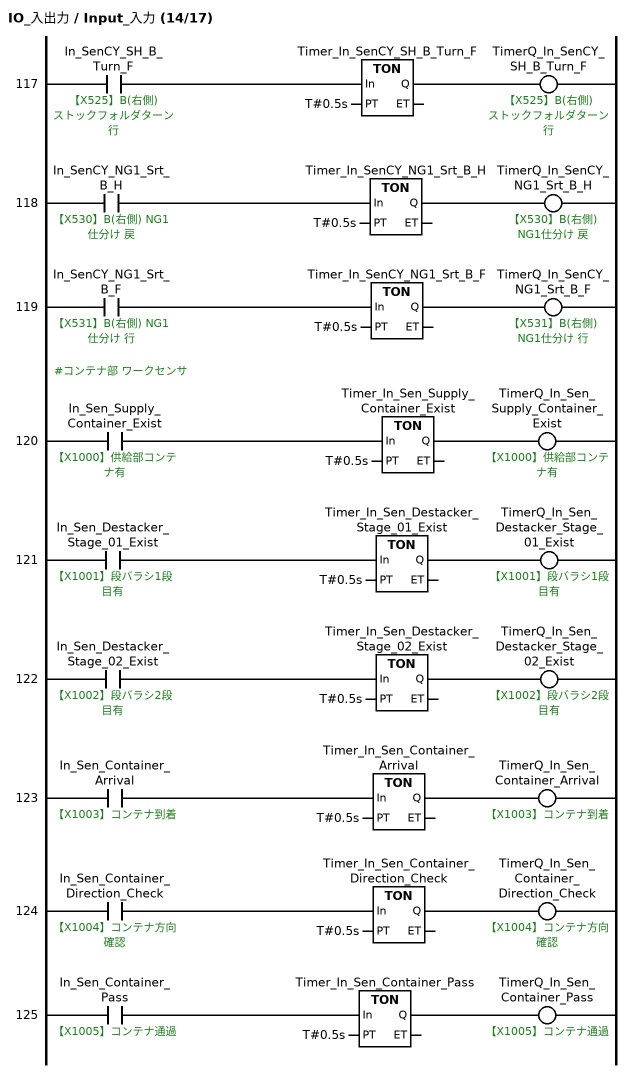
(* [picture p188: IO_入出力 / Input_入力, rungs 117-125] *)
(* Rung 117 *)
Timer_In_SenCY_SH_B_Turn_F(In := In_SenCY_SH_B_Turn_F, PT := T#0.5s);
TimerQ_In_SenCY_SH_B_Turn_F := Timer_In_SenCY_SH_B_Turn_F.Q;
(* Rung 118 *)
Timer_In_SenCY_NG1_Srt_B_H(In := In_SenCY_NG1_Srt_B_H, PT := T#0.5s);
TimerQ_In_SenCY_NG1_Srt_B_H := Timer_In_SenCY_NG1_Srt_B_H.Q;
(* Rung 119 *)
Timer_In_SenCY_NG1_Srt_B_F(In := In_SenCY_NG1_Srt_B_F, PT := T#0.5s);
TimerQ_In_SenCY_NG1_Srt_B_F := Timer_In_SenCY_NG1_Srt_B_F.Q;
(* Rung 120: #コンテナ部 ワークセンサ *)
Timer_In_Sen_Supply_Container_Exist(In := In_Sen_Supply_Container_Exist, PT := T#0.5s);
TimerQ_In_Sen_Supply_Container_Exist := Timer_In_Sen_Supply_Container_Exist.Q;
(* Rung 121 *)
Timer_In_Sen_Destacker_Stage_01_Exist(In := In_Sen_Destacker_Stage_01_Exist, PT := T#0.5s);
TimerQ_In_Sen_Destacker_Stage_01_Exist := Timer_In_Sen_Destacker_Stage_01_Exist.Q;
(* Rung 122 *)
Timer_In_Sen_Destacker_Stage_02_Exist(In := In_Sen_Destacker_Stage_02_Exist, PT := T#0.5s);
TimerQ_In_Sen_Destacker_Stage_02_Exist := Timer_In_Sen_Destacker_Stage_02_Exist.Q;
(* Rung 123 *)
Timer_In_Sen_Container_Arrival(In := In_Sen_Container_Arrival, PT := T#0.5s);
TimerQ_In_Sen_Container_Arrival := Timer_In_Sen_Container_Arrival.Q;
(* Rung 124 *)
Timer_In_Sen_Container_Direction_Check(In := In_Sen_Container_Direction_Check, PT := T#0.5s);
TimerQ_In_Sen_Container_Direction_Check := Timer_In_Sen_Container_Direction_Check.Q;
(* Rung 125 *)
Timer_In_Sen_Container_Pass(In := In_Sen_Container_Pass, PT := T#0.5s);
TimerQ_In_Sen_Container_Pass := Timer_In_Sen_Container_Pass.Q;

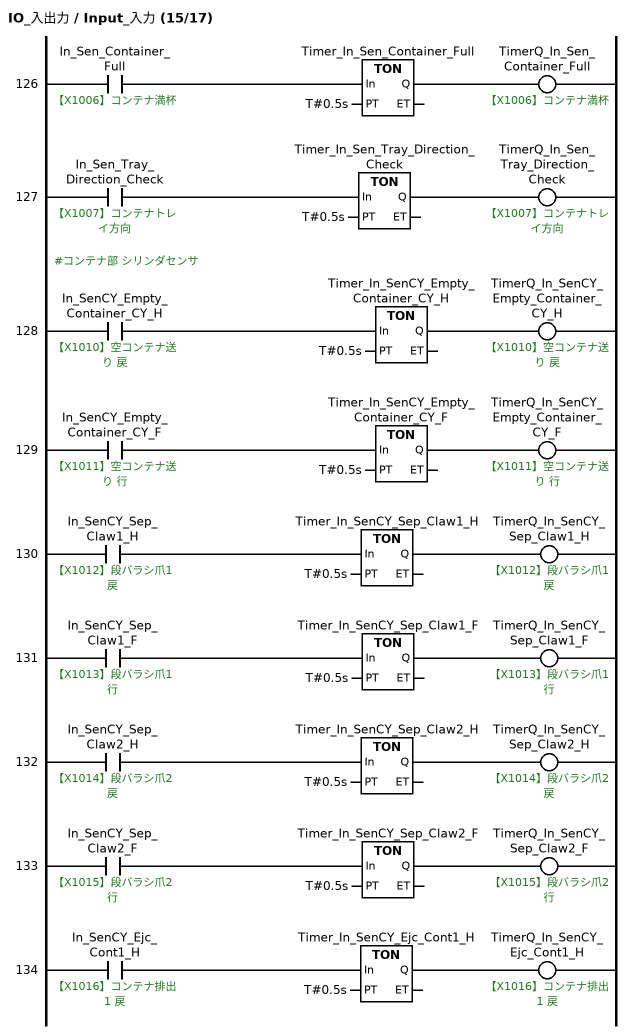
(* Rung 126 *)
Timer_In_Sen_Container_Full(In := In_Sen_Container_Full, PT := T#0.5s);
TimerQ_In_Sen_Container_Full := Timer_In_Sen_Container_Full.Q;
(* Rung 127 *)
Timer_In_Sen_Tray_Direction_Check(In := In_Sen_Tray_Direction_Check, PT := T#0.5s);
TimerQ_In_Sen_Tray_Direction_Check := Timer_In_Sen_Tray_Direction_Check.Q;
(* Rung 128: #コンテナ部 シリンダセンサ *)
Timer_In_SenCY_Empty_Container_CY_H(In := In_SenCY_Empty_Container_CY_H, PT := T#0.5s);
TimerQ_In_SenCY_Empty_Container_CY_H := Timer_In_SenCY_Empty_Container_CY_H.Q;
(* Rung 129 *)
Timer_In_SenCY_Empty_Container_CY_F(In := In_SenCY_Empty_Container_CY_F, PT := T#0.5s);
TimerQ_In_SenCY_Empty_Container_CY_F := Timer_In_SenCY_Empty_Container_CY_F.Q;
(* Rung 130 *)
Timer_In_SenCY_Sep_Claw1_H(In := In_SenCY_Sep_Claw1_H, PT := T#0.5s);
TimerQ_In_SenCY_Sep_Claw1_H := Timer_In_SenCY_Sep_Claw1_H.Q;
(* Rung 131 *)
Timer_In_SenCY_Sep_Claw1_F(In := In_SenCY_Sep_Claw1_F, PT := T#0.5s);
TimerQ_In_SenCY_Sep_Claw1_F := Timer_In_SenCY_Sep_Claw1_F.Q;
(* Rung 132 *)
Timer_In_SenCY_Sep_Claw2_H(In := In_SenCY_Sep_Claw2_H, PT := T#0.5s);
TimerQ_In_SenCY_Sep_Claw2_H := Timer_In_SenCY_Sep_Claw2_H.Q;
(* Rung 133 *)
Timer_In_SenCY_Sep_Claw2_F(In := In_SenCY_Sep_Claw2_F, PT := T#0.5s);
TimerQ_In_SenCY_Sep_Claw2_F := Timer_In_SenCY_Sep_Claw2_F.Q;
(* Rung 134 *)
Timer_In_SenCY_Ejc_Cont1_H(In := In_SenCY_Ejc_Cont1_H, PT := T#0.5s);
TimerQ_In_SenCY_Ejc_Cont1_H := Timer_In_SenCY_Ejc_Cont1_H.Q;

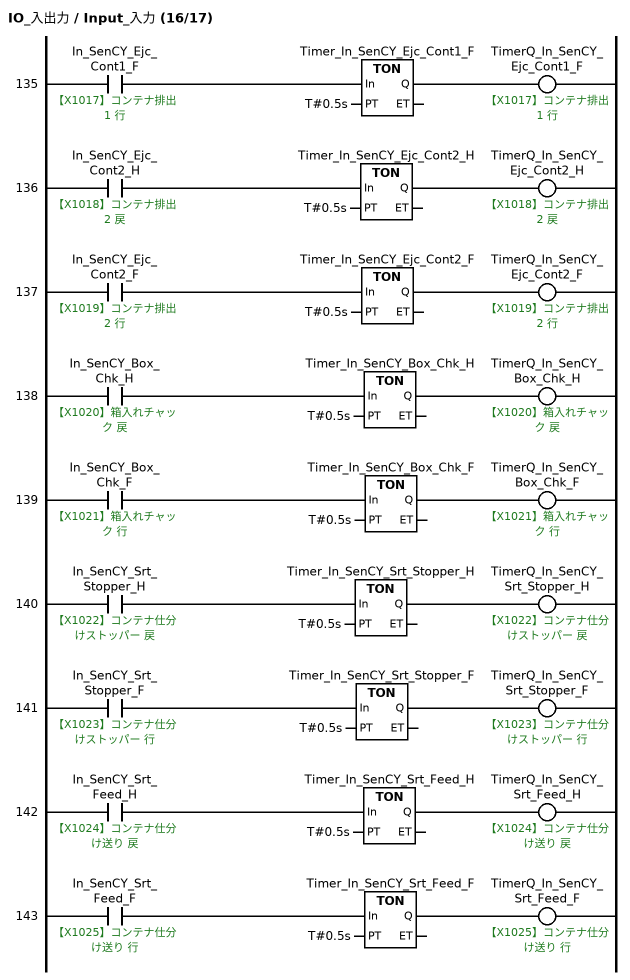
(* Rung 135 *)
Timer_In_SenCY_Ejc_Cont1_F(In := In_SenCY_Ejc_Cont1_F, PT := T#0.5s);
TimerQ_In_SenCY_Ejc_Cont1_F := Timer_In_SenCY_Ejc_Cont1_F.Q;
(* Rung 136 *)
Timer_In_SenCY_Ejc_Cont2_H(In := In_SenCY_Ejc_Cont2_H, PT := T#0.5s);
TimerQ_In_SenCY_Ejc_Cont2_H := Timer_In_SenCY_Ejc_Cont2_H.Q;
(* Rung 137 *)
Timer_In_SenCY_Ejc_Cont2_F(In := In_SenCY_Ejc_Cont2_F, PT := T#0.5s);
TimerQ_In_SenCY_Ejc_Cont2_F := Timer_In_SenCY_Ejc_Cont2_F.Q;
(* Rung 138 *)
Timer_In_SenCY_Box_Chk_H(In := In_SenCY_Box_Chk_H, PT := T#0.5s);
TimerQ_In_SenCY_Box_Chk_H := Timer_In_SenCY_Box_Chk_H.Q;
(* Rung 139 *)
Timer_In_SenCY_Box_Chk_F(In := In_SenCY_Box_Chk_F, PT := T#0.5s);
TimerQ_In_SenCY_Box_Chk_F := Timer_In_SenCY_Box_Chk_F.Q;
(* Rung 140 *)
Timer_In_SenCY_Srt_Stopper_H(In := In_SenCY_Srt_Stopper_H, PT := T#0.5s);
TimerQ_In_SenCY_Srt_Stopper_H := Timer_In_SenCY_Srt_Stopper_H.Q;
(* Rung 141 *)
Timer_In_SenCY_Srt_Stopper_F(In := In_SenCY_Srt_Stopper_F, PT := T#0.5s);
TimerQ_In_SenCY_Srt_Stopper_F := Timer_In_SenCY_Srt_Stopper_F.Q;
(* Rung 142 *)
Timer_In_SenCY_Srt_Feed_H(In := In_SenCY_Srt_Feed_H, PT := T#0.5s);
TimerQ_In_SenCY_Srt_Feed_H := Timer_In_SenCY_Srt_Feed_H.Q;
(* Rung 143 *)
Timer_In_SenCY_Srt_Feed_F(In := In_SenCY_Srt_Feed_F, PT := T#0.5s);
TimerQ_In_SenCY_Srt_Feed_F := Timer_In_SenCY_Srt_Feed_F.Q;

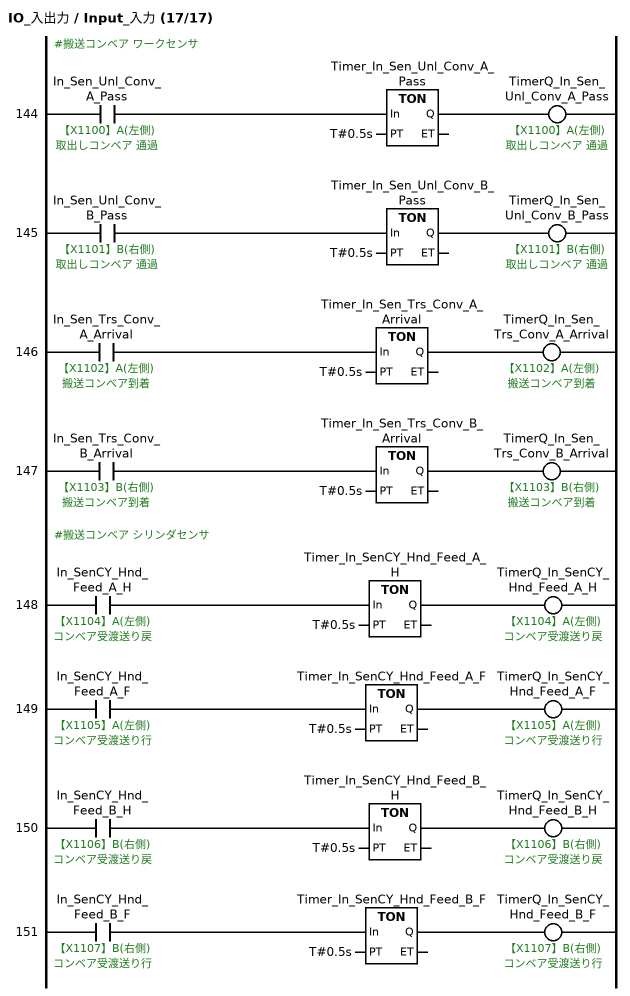
(* Rung 144: #搬送コンベア ワークセンサ *)
Timer_In_Sen_Unl_Conv_A_Pass(In := In_Sen_Unl_Conv_A_Pass, PT := T#0.5s);
TimerQ_In_Sen_Unl_Conv_A_Pass := Timer_In_Sen_Unl_Conv_A_Pass.Q;
(* Rung 145 *)
Timer_In_Sen_Unl_Conv_B_Pass(In := In_Sen_Unl_Conv_B_Pass, PT := T#0.5s);
TimerQ_In_Sen_Unl_Conv_B_Pass := Timer_In_Sen_Unl_Conv_B_Pass.Q;
(* Rung 146 *)
Timer_In_Sen_Trs_Conv_A_Arrival(In := In_Sen_Trs_Conv_A_Arrival, PT := T#0.5s);
TimerQ_In_Sen_Trs_Conv_A_Arrival := Timer_In_Sen_Trs_Conv_A_Arrival.Q;
(* Rung 147 *)
Timer_In_Sen_Trs_Conv_B_Arrival(In := In_Sen_Trs_Conv_B_Arrival, PT := T#0.5s);
TimerQ_In_Sen_Trs_Conv_B_Arrival := Timer_In_Sen_Trs_Conv_B_Arrival.Q;
(* Rung 148: #搬送コンベア シリンダセンサ *)
Timer_In_SenCY_Hnd_Feed_A_H(In := In_SenCY_Hnd_Feed_A_H, PT := T#0.5s);
TimerQ_In_SenCY_Hnd_Feed_A_H := Timer_In_SenCY_Hnd_Feed_A_H.Q;
(* Rung 149 *)
Timer_In_SenCY_Hnd_Feed_A_F(In := In_SenCY_Hnd_Feed_A_F, PT := T#0.5s);
TimerQ_In_SenCY_Hnd_Feed_A_F := Timer_In_SenCY_Hnd_Feed_A_F.Q;
(* Rung 150 *)
Timer_In_SenCY_Hnd_Feed_B_H(In := In_SenCY_Hnd_Feed_B_H, PT := T#0.5s);
TimerQ_In_SenCY_Hnd_Feed_B_H := Timer_In_SenCY_Hnd_Feed_B_H.Q;
(* Rung 151 *)
Timer_In_SenCY_Hnd_Feed_B_F(In := In_SenCY_Hnd_Feed_B_F, PT := T#0.5s);
TimerQ_In_SenCY_Hnd_Feed_B_F := Timer_In_SenCY_Hnd_Feed_B_F.Q;

(* Section Output_出力: ladder, written here as Structured Text *)

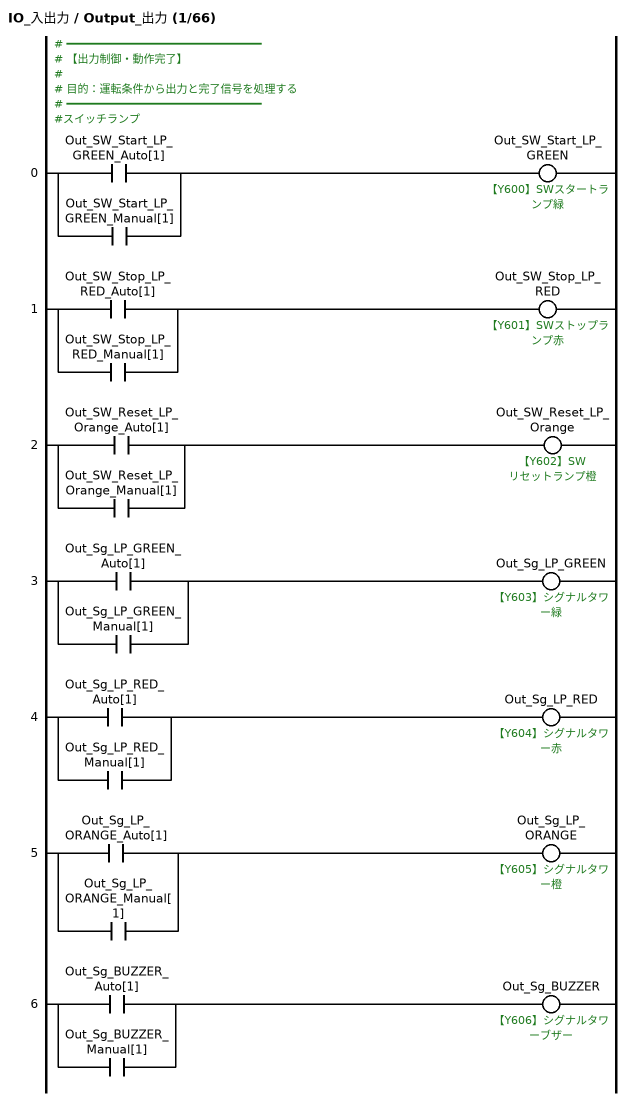
(* Rung 0: # ━━━━━━━━━━━━━━━━━━━━━━━━━━━━━━ / # 【出力制御・動作完了】 / # / # 目的：運転条件から出力と完了信号を処理する / # ━━━━━━━━━━━━━━━━━━━━━━━━━━━━━━ / #スイッチランプ *)
Out_SW_Start_LP_GREEN := Out_SW_Start_LP_GREEN_Auto[1] OR Out_SW_Start_LP_GREEN_Manual[1];
(* Rung 1 *)
Out_SW_Stop_LP_RED := Out_SW_Stop_LP_RED_Auto[1] OR Out_SW_Stop_LP_RED_Manual[1];
(* Rung 2 *)
Out_SW_Reset_LP_Orange := Out_SW_Reset_LP_Orange_Auto[1] OR Out_SW_Reset_LP_Orange_Manual[1];
(* Rung 3 *)
Out_Sg_LP_GREEN := Out_Sg_LP_GREEN_Auto[1] OR Out_Sg_LP_GREEN_Manual[1];
(* Rung 4 *)
Out_Sg_LP_RED := Out_Sg_LP_RED_Auto[1] OR Out_Sg_LP_RED_Manual[1];
(* Rung 5 *)
Out_Sg_LP_ORANGE := Out_Sg_LP_ORANGE_Auto[1] OR Out_Sg_LP_ORANGE_Manual[1];
(* Rung 6 *)
Out_Sg_BUZZER := Out_Sg_BUZZER_Auto[1] OR Out_Sg_BUZZER_Manual[1];

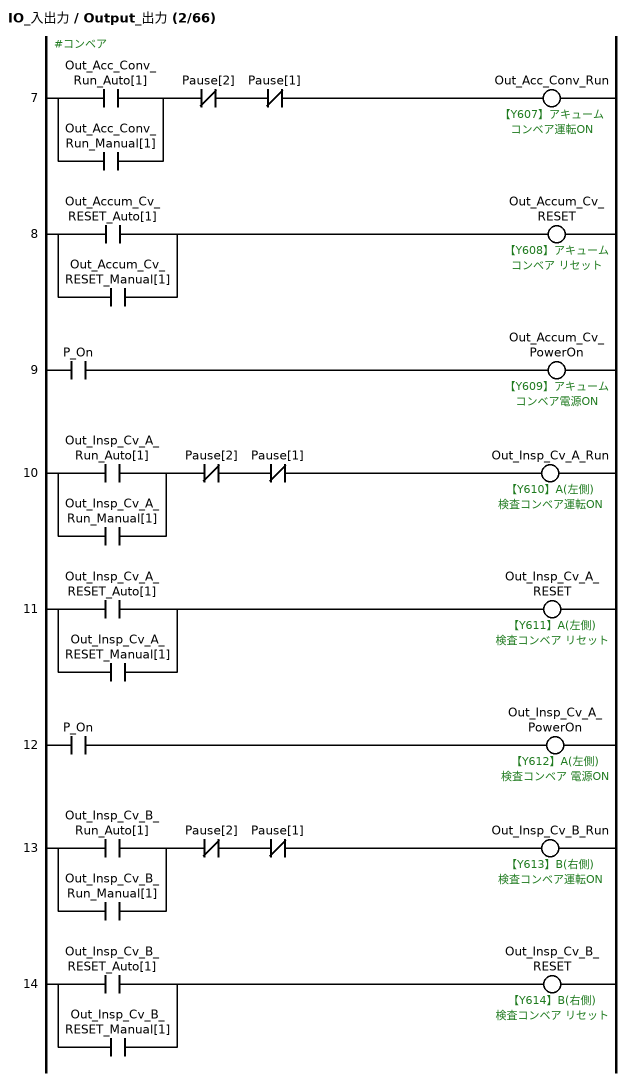
(* Rung 7: #コンベア *)
Out_Acc_Conv_Run := (Out_Acc_Conv_Run_Auto[1] OR Out_Acc_Conv_Run_Manual[1]) AND NOT Pause[2] AND NOT Pause[1];
(* Rung 8 *)
Out_Accum_Cv_RESET := Out_Accum_Cv_RESET_Auto[1] OR Out_Accum_Cv_RESET_Manual[1];
(* Rung 9 *)
Out_Accum_Cv_PowerOn := P_On;
(* Rung 10 *)
Out_Insp_Cv_A_Run := (Out_Insp_Cv_A_Run_Auto[1] OR Out_Insp_Cv_A_Run_Manual[1]) AND NOT Pause[2] AND NOT Pause[1];
(* Rung 11 *)
Out_Insp_Cv_A_RESET := Out_Insp_Cv_A_RESET_Auto[1] OR Out_Insp_Cv_A_RESET_Manual[1];
(* Rung 12 *)
Out_Insp_Cv_A_PowerOn := P_On;
(* Rung 13 *)
Out_Insp_Cv_B_Run := (Out_Insp_Cv_B_Run_Auto[1] OR Out_Insp_Cv_B_Run_Manual[1]) AND NOT Pause[2] AND NOT Pause[1];
(* Rung 14 *)
Out_Insp_Cv_B_RESET := Out_Insp_Cv_B_RESET_Auto[1] OR Out_Insp_Cv_B_RESET_Manual[1];

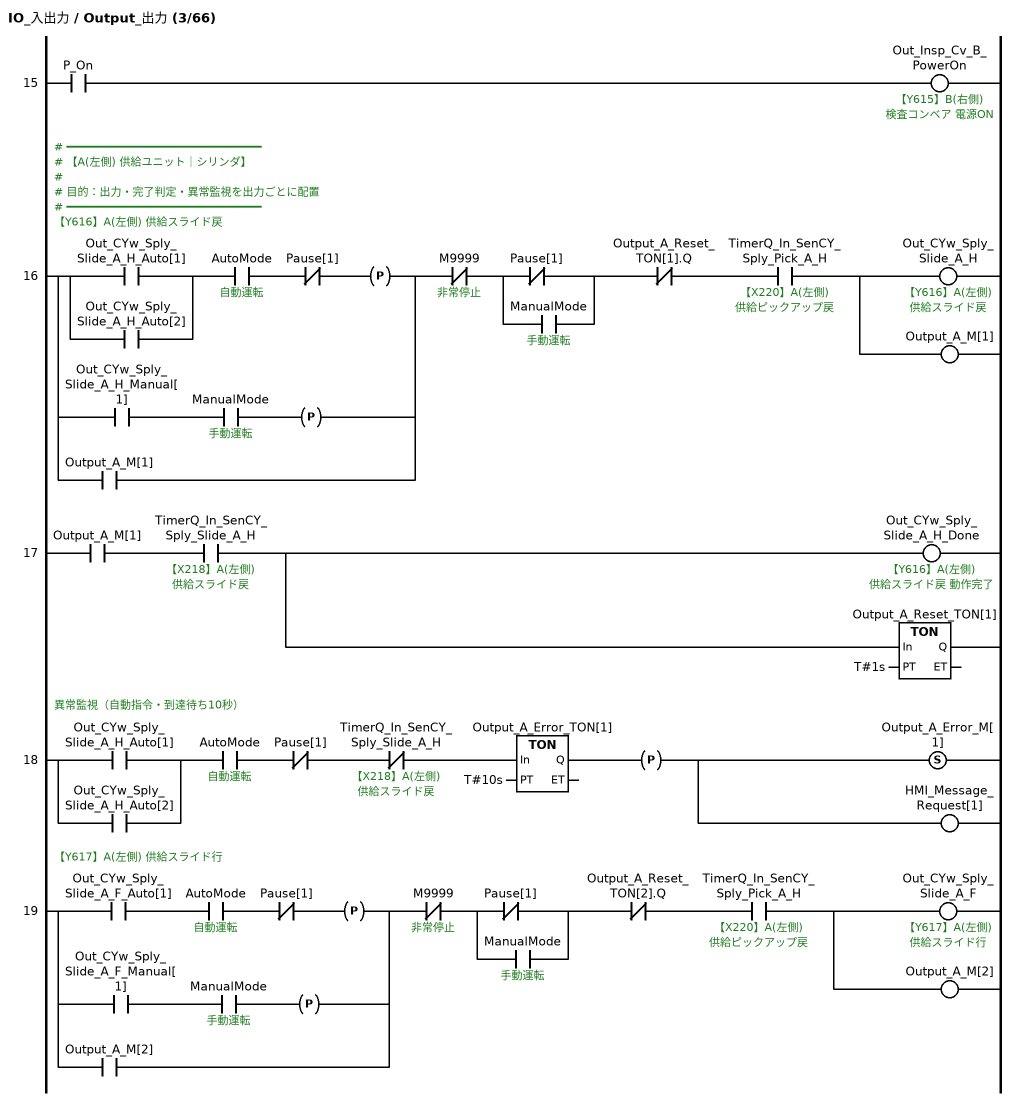
(* Rung 15 *)
Out_Insp_Cv_B_PowerOn := P_On;
(* Rung 16: # ━━━━━━━━━━━━━━━━━━━━━━━━━━━━━━ / # 【A(左側) 供給ユニット｜シリンダ】 / # / # 目的：出力・完了判定・異常監視を出力ごとに配置 / # ━━━━━━━━━━━━━━━━━━━━━━━━━━━━━━ / 【Y616】A(左側) 供給スライド戻 *)
_e1(CLK := (Out_CYw_Sply_Slide_A_H_Auto[1] OR Out_CYw_Sply_Slide_A_H_Auto[2]) AND AutoMode AND NOT Pause[1]);
_e2(CLK := Out_CYw_Sply_Slide_A_H_Manual[1] AND ManualMode);
_p3 := (_e1.Q OR _e2.Q OR Output_A_M[1]) AND NOT M9999 AND (NOT Pause[1] OR ManualMode) AND NOT Output_A_Reset_TON[1].Q AND TimerQ_In_SenCY_Sply_Pick_A_H;
Out_CYw_Sply_Slide_A_H := _p3;
Output_A_M[1] := _p3;
(* Rung 17 *)
Out_CYw_Sply_Slide_A_H_Done := Output_A_M[1] AND TimerQ_In_SenCY_Sply_Slide_A_H;
Output_A_Reset_TON[1](In := Output_A_M[1] AND TimerQ_In_SenCY_Sply_Slide_A_H, PT := T#1s);
(* Rung 18: 異常監視（自動指令・到達待ち10秒） *)
Output_A_Error_TON[1](In := (Out_CYw_Sply_Slide_A_H_Auto[1] OR Out_CYw_Sply_Slide_A_H_Auto[2]) AND AutoMode AND NOT Pause[1] AND NOT TimerQ_In_SenCY_Sply_Slide_A_H, PT := T#10s);
_e4(CLK := Output_A_Error_TON[1].Q);
IF _e4.Q THEN Output_A_Error_M[1] := TRUE; END_IF;
HMI_Message_Request[1] := _e4.Q;
(* Rung 19: 【Y617】A(左側) 供給スライド行 *)
_e5(CLK := Out_CYw_Sply_Slide_A_F_Auto[1] AND AutoMode AND NOT Pause[1]);
_e6(CLK := Out_CYw_Sply_Slide_A_F_Manual[1] AND ManualMode);
_p7 := (_e5.Q OR _e6.Q OR Output_A_M[2]) AND NOT M9999 AND (NOT Pause[1] OR ManualMode) AND NOT Output_A_Reset_TON[2].Q AND TimerQ_In_SenCY_Sply_Pick_A_H;
Out_CYw_Sply_Slide_A_F := _p7;
Output_A_M[2] := _p7;

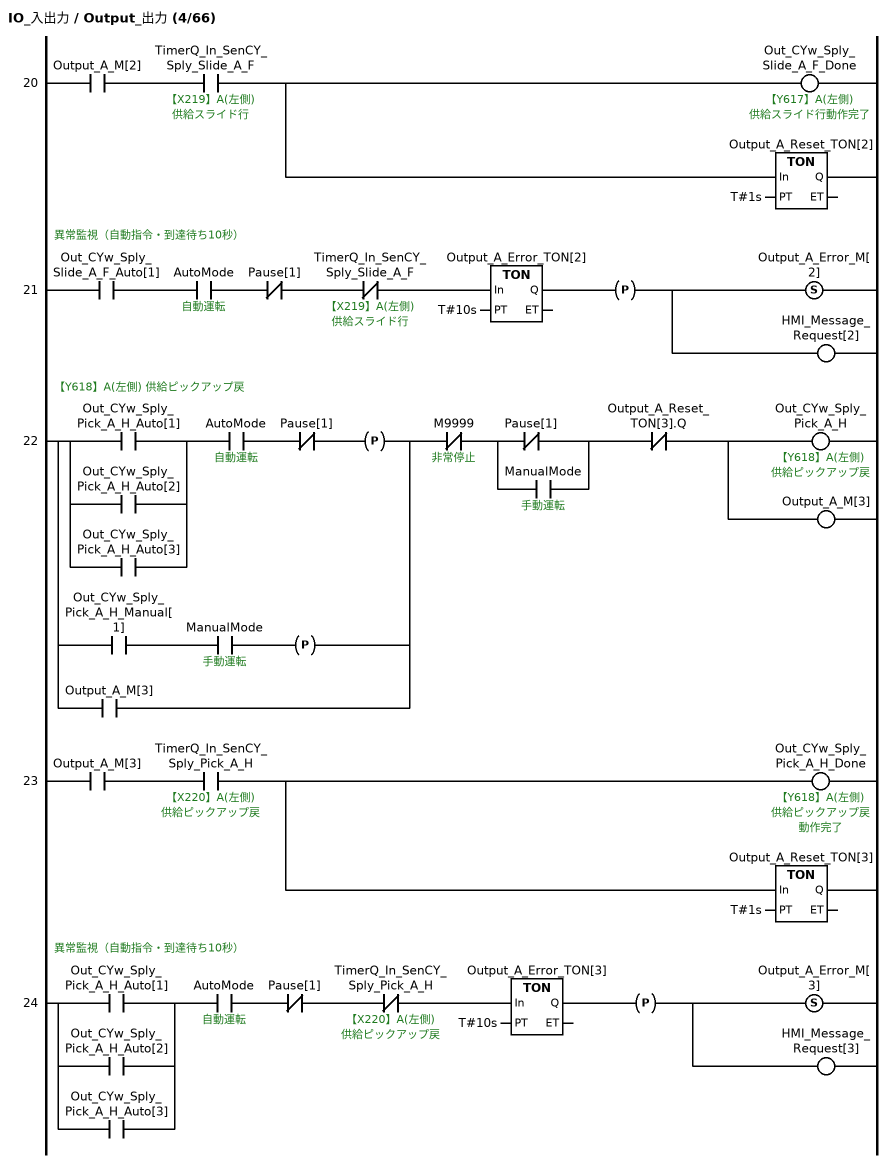
(* Rung 20 *)
Out_CYw_Sply_Slide_A_F_Done := Output_A_M[2] AND TimerQ_In_SenCY_Sply_Slide_A_F;
Output_A_Reset_TON[2](In := Output_A_M[2] AND TimerQ_In_SenCY_Sply_Slide_A_F, PT := T#1s);
(* Rung 21: 異常監視（自動指令・到達待ち10秒） *)
Output_A_Error_TON[2](In := Out_CYw_Sply_Slide_A_F_Auto[1] AND AutoMode AND NOT Pause[1] AND NOT TimerQ_In_SenCY_Sply_Slide_A_F, PT := T#10s);
_e8(CLK := Output_A_Error_TON[2].Q);
IF _e8.Q THEN Output_A_Error_M[2] := TRUE; END_IF;
HMI_Message_Request[2] := _e8.Q;
(* Rung 22: 【Y618】A(左側) 供給ピックアップ戻 *)
_e9(CLK := (Out_CYw_Sply_Pick_A_H_Auto[1] OR Out_CYw_Sply_Pick_A_H_Auto[2] OR Out_CYw_Sply_Pick_A_H_Auto[3]) AND AutoMode AND NOT Pause[1]);
_e10(CLK := Out_CYw_Sply_Pick_A_H_Manual[1] AND ManualMode);
_p11 := (_e9.Q OR _e10.Q OR Output_A_M[3]) AND NOT M9999 AND (NOT Pause[1] OR ManualMode) AND NOT Output_A_Reset_TON[3].Q;
Out_CYw_Sply_Pick_A_H := _p11;
Output_A_M[3] := _p11;
(* Rung 23 *)
Out_CYw_Sply_Pick_A_H_Done := Output_A_M[3] AND TimerQ_In_SenCY_Sply_Pick_A_H;
Output_A_Reset_TON[3](In := Output_A_M[3] AND TimerQ_In_SenCY_Sply_Pick_A_H, PT := T#1s);
(* Rung 24: 異常監視（自動指令・到達待ち10秒） *)
Output_A_Error_TON[3](In := (Out_CYw_Sply_Pick_A_H_Auto[1] OR Out_CYw_Sply_Pick_A_H_Auto[2] OR Out_CYw_Sply_Pick_A_H_Auto[3]) AND AutoMode AND NOT Pause[1] AND NOT TimerQ_In_SenCY_Sply_Pick_A_H, PT := T#10s);
_e12(CLK := Output_A_Error_TON[3].Q);
IF _e12.Q THEN Output_A_Error_M[3] := TRUE; END_IF;
HMI_Message_Request[3] := _e12.Q;

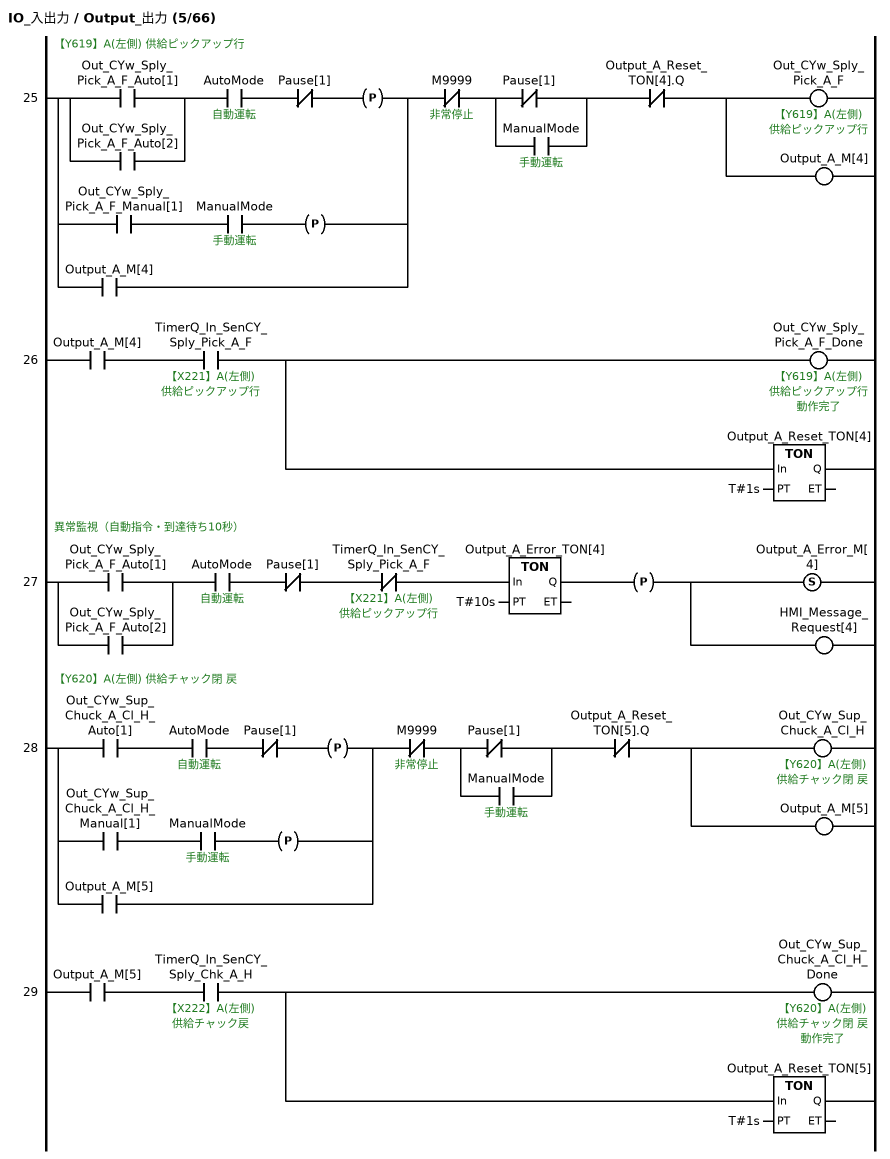
(* Rung 25: 【Y619】A(左側) 供給ピックアップ行 *)
_e13(CLK := (Out_CYw_Sply_Pick_A_F_Auto[1] OR Out_CYw_Sply_Pick_A_F_Auto[2]) AND AutoMode AND NOT Pause[1]);
_e14(CLK := Out_CYw_Sply_Pick_A_F_Manual[1] AND ManualMode);
_p15 := (_e13.Q OR _e14.Q OR Output_A_M[4]) AND NOT M9999 AND (NOT Pause[1] OR ManualMode) AND NOT Output_A_Reset_TON[4].Q;
Out_CYw_Sply_Pick_A_F := _p15;
Output_A_M[4] := _p15;
(* Rung 26 *)
Out_CYw_Sply_Pick_A_F_Done := Output_A_M[4] AND TimerQ_In_SenCY_Sply_Pick_A_F;
Output_A_Reset_TON[4](In := Output_A_M[4] AND TimerQ_In_SenCY_Sply_Pick_A_F, PT := T#1s);
(* Rung 27: 異常監視（自動指令・到達待ち10秒） *)
Output_A_Error_TON[4](In := (Out_CYw_Sply_Pick_A_F_Auto[1] OR Out_CYw_Sply_Pick_A_F_Auto[2]) AND AutoMode AND NOT Pause[1] AND NOT TimerQ_In_SenCY_Sply_Pick_A_F, PT := T#10s);
_e16(CLK := Output_A_Error_TON[4].Q);
IF _e16.Q THEN Output_A_Error_M[4] := TRUE; END_IF;
HMI_Message_Request[4] := _e16.Q;
(* Rung 28: 【Y620】A(左側) 供給チャック閉 戻 *)
_e17(CLK := Out_CYw_Sup_Chuck_A_Cl_H_Auto[1] AND AutoMode AND NOT Pause[1]);
_e18(CLK := Out_CYw_Sup_Chuck_A_Cl_H_Manual[1] AND ManualMode);
_p19 := (_e17.Q OR _e18.Q OR Output_A_M[5]) AND NOT M9999 AND (NOT Pause[1] OR ManualMode) AND NOT Output_A_Reset_TON[5].Q;
Out_CYw_Sup_Chuck_A_Cl_H := _p19;
Output_A_M[5] := _p19;
(* Rung 29 *)
Out_CYw_Sup_Chuck_A_Cl_H_Done := Output_A_M[5] AND TimerQ_In_SenCY_Sply_Chk_A_H;
Output_A_Reset_TON[5](In := Output_A_M[5] AND TimerQ_In_SenCY_Sply_Chk_A_H, PT := T#1s);

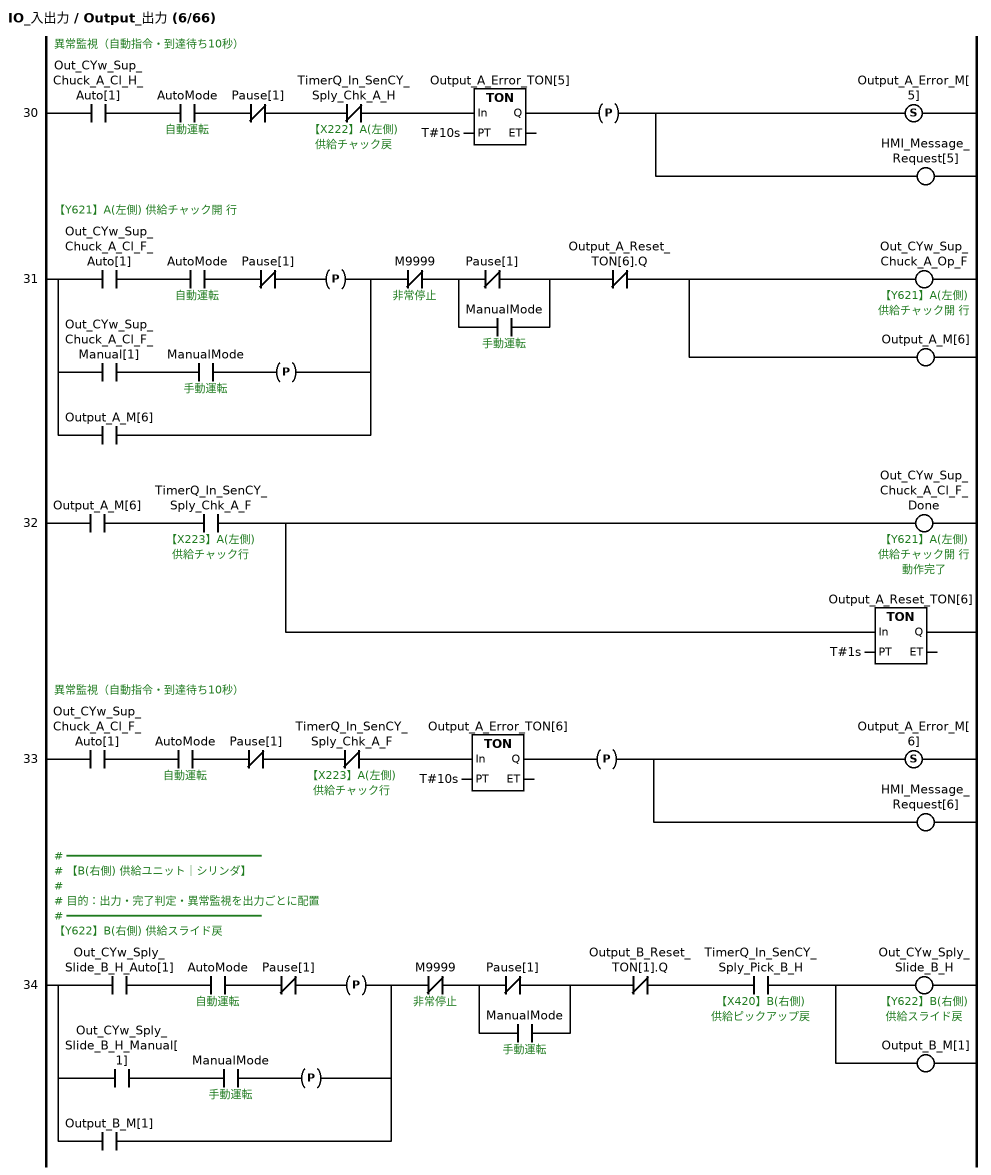
(* Rung 30: 異常監視（自動指令・到達待ち10秒） *)
Output_A_Error_TON[5](In := Out_CYw_Sup_Chuck_A_Cl_H_Auto[1] AND AutoMode AND NOT Pause[1] AND NOT TimerQ_In_SenCY_Sply_Chk_A_H, PT := T#10s);
_e20(CLK := Output_A_Error_TON[5].Q);
IF _e20.Q THEN Output_A_Error_M[5] := TRUE; END_IF;
HMI_Message_Request[5] := _e20.Q;
(* Rung 31: 【Y621】A(左側) 供給チャック開 行 *)
_e21(CLK := Out_CYw_Sup_Chuck_A_Cl_F_Auto[1] AND AutoMode AND NOT Pause[1]);
_e22(CLK := Out_CYw_Sup_Chuck_A_Cl_F_Manual[1] AND ManualMode);
_p23 := (_e21.Q OR _e22.Q OR Output_A_M[6]) AND NOT M9999 AND (NOT Pause[1] OR ManualMode) AND NOT Output_A_Reset_TON[6].Q;
Out_CYw_Sup_Chuck_A_Op_F := _p23;
Output_A_M[6] := _p23;
(* Rung 32 *)
Out_CYw_Sup_Chuck_A_Cl_F_Done := Output_A_M[6] AND TimerQ_In_SenCY_Sply_Chk_A_F;
Output_A_Reset_TON[6](In := Output_A_M[6] AND TimerQ_In_SenCY_Sply_Chk_A_F, PT := T#1s);
(* Rung 33: 異常監視（自動指令・到達待ち10秒） *)
Output_A_Error_TON[6](In := Out_CYw_Sup_Chuck_A_Cl_F_Auto[1] AND AutoMode AND NOT Pause[1] AND NOT TimerQ_In_SenCY_Sply_Chk_A_F, PT := T#10s);
_e24(CLK := Output_A_Error_TON[6].Q);
IF _e24.Q THEN Output_A_Error_M[6] := TRUE; END_IF;
HMI_Message_Request[6] := _e24.Q;
(* Rung 34: # ━━━━━━━━━━━━━━━━━━━━━━━━━━━━━━ / # 【B(右側) 供給ユニット｜シリンダ】 / # / # 目的：出力・完了判定・異常監視を出力ごとに配置 / # ━━━━━━━━━━━━━━━━━━━━━━━━━━━━━━ / 【Y622】B(右側) 供給スライド戻 *)
_e25(CLK := Out_CYw_Sply_Slide_B_H_Auto[1] AND AutoMode AND NOT Pause[1]);
_e26(CLK := Out_CYw_Sply_Slide_B_H_Manual[1] AND ManualMode);
_p27 := (_e25.Q OR _e26.Q OR Output_B_M[1]) AND NOT M9999 AND (NOT Pause[1] OR ManualMode) AND NOT Output_B_Reset_TON[1].Q AND TimerQ_In_SenCY_Sply_Pick_B_H;
Out_CYw_Sply_Slide_B_H := _p27;
Output_B_M[1] := _p27;

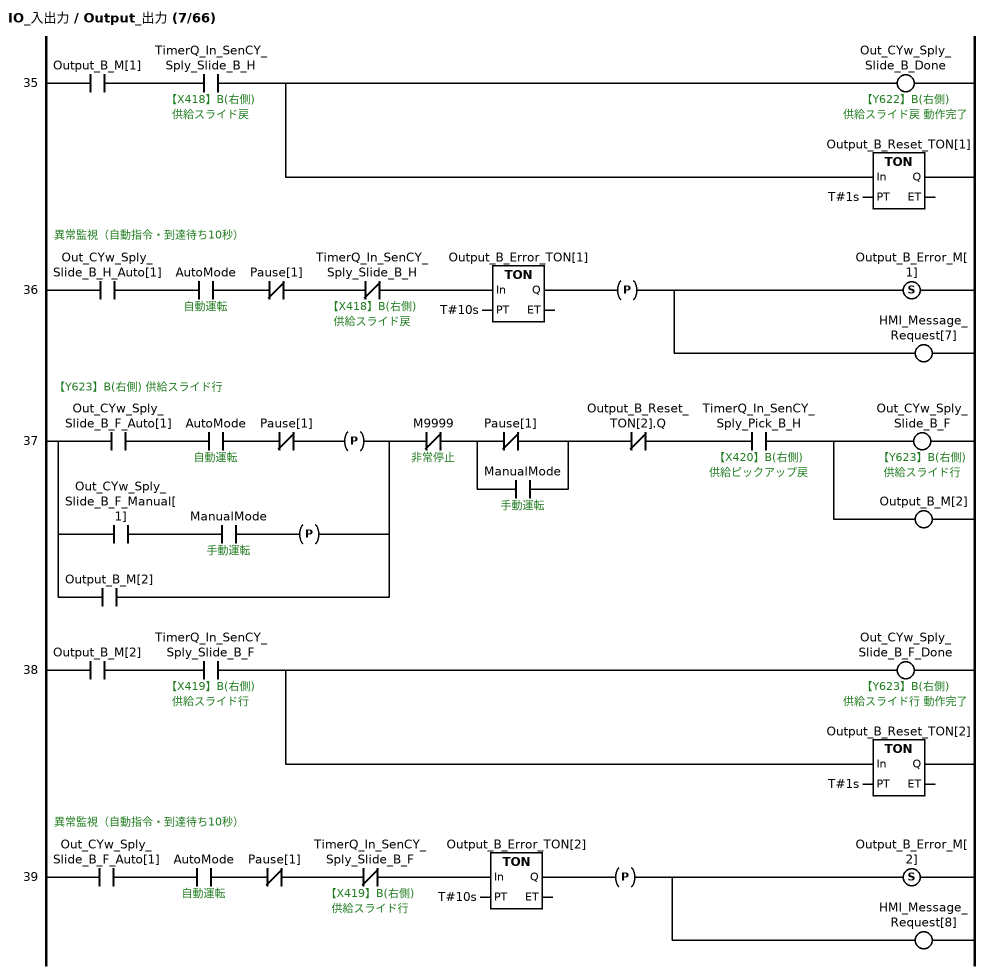
(* Rung 35 *)
Out_CYw_Sply_Slide_B_Done := Output_B_M[1] AND TimerQ_In_SenCY_Sply_Slide_B_H;
Output_B_Reset_TON[1](In := Output_B_M[1] AND TimerQ_In_SenCY_Sply_Slide_B_H, PT := T#1s);
(* Rung 36: 異常監視（自動指令・到達待ち10秒） *)
Output_B_Error_TON[1](In := Out_CYw_Sply_Slide_B_H_Auto[1] AND AutoMode AND NOT Pause[1] AND NOT TimerQ_In_SenCY_Sply_Slide_B_H, PT := T#10s);
_e28(CLK := Output_B_Error_TON[1].Q);
IF _e28.Q THEN Output_B_Error_M[1] := TRUE; END_IF;
HMI_Message_Request[7] := _e28.Q;
(* Rung 37: 【Y623】B(右側) 供給スライド行 *)
_e29(CLK := Out_CYw_Sply_Slide_B_F_Auto[1] AND AutoMode AND NOT Pause[1]);
_e30(CLK := Out_CYw_Sply_Slide_B_F_Manual[1] AND ManualMode);
_p31 := (_e29.Q OR _e30.Q OR Output_B_M[2]) AND NOT M9999 AND (NOT Pause[1] OR ManualMode) AND NOT Output_B_Reset_TON[2].Q AND TimerQ_In_SenCY_Sply_Pick_B_H;
Out_CYw_Sply_Slide_B_F := _p31;
Output_B_M[2] := _p31;
(* Rung 38 *)
Out_CYw_Sply_Slide_B_F_Done := Output_B_M[2] AND TimerQ_In_SenCY_Sply_Slide_B_F;
Output_B_Reset_TON[2](In := Output_B_M[2] AND TimerQ_In_SenCY_Sply_Slide_B_F, PT := T#1s);
(* Rung 39: 異常監視（自動指令・到達待ち10秒） *)
Output_B_Error_TON[2](In := Out_CYw_Sply_Slide_B_F_Auto[1] AND AutoMode AND NOT Pause[1] AND NOT TimerQ_In_SenCY_Sply_Slide_B_F, PT := T#10s);
_e32(CLK := Output_B_Error_TON[2].Q);
IF _e32.Q THEN Output_B_Error_M[2] := TRUE; END_IF;
HMI_Message_Request[8] := _e32.Q;

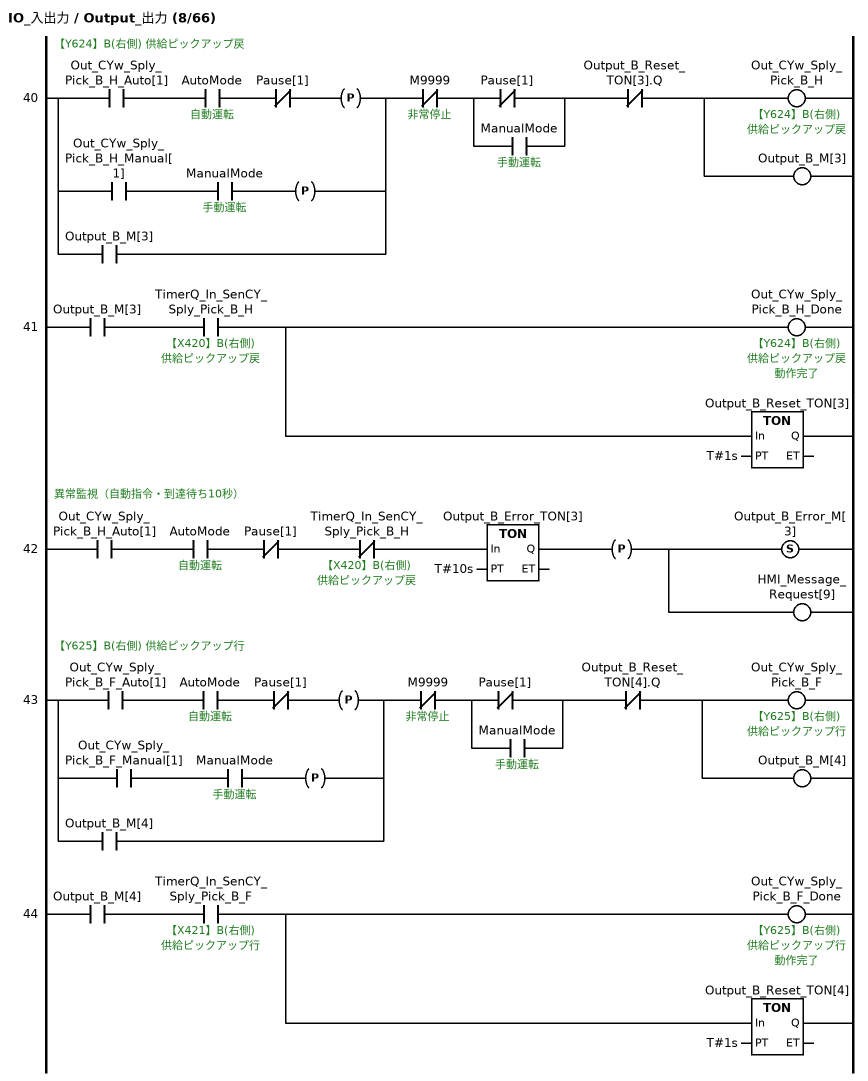
(* Rung 40: 【Y624】B(右側) 供給ピックアップ戻 *)
_e33(CLK := Out_CYw_Sply_Pick_B_H_Auto[1] AND AutoMode AND NOT Pause[1]);
_e34(CLK := Out_CYw_Sply_Pick_B_H_Manual[1] AND ManualMode);
_p35 := (_e33.Q OR _e34.Q OR Output_B_M[3]) AND NOT M9999 AND (NOT Pause[1] OR ManualMode) AND NOT Output_B_Reset_TON[3].Q;
Out_CYw_Sply_Pick_B_H := _p35;
Output_B_M[3] := _p35;
(* Rung 41 *)
Out_CYw_Sply_Pick_B_H_Done := Output_B_M[3] AND TimerQ_In_SenCY_Sply_Pick_B_H;
Output_B_Reset_TON[3](In := Output_B_M[3] AND TimerQ_In_SenCY_Sply_Pick_B_H, PT := T#1s);
(* Rung 42: 異常監視（自動指令・到達待ち10秒） *)
Output_B_Error_TON[3](In := Out_CYw_Sply_Pick_B_H_Auto[1] AND AutoMode AND NOT Pause[1] AND NOT TimerQ_In_SenCY_Sply_Pick_B_H, PT := T#10s);
_e36(CLK := Output_B_Error_TON[3].Q);
IF _e36.Q THEN Output_B_Error_M[3] := TRUE; END_IF;
HMI_Message_Request[9] := _e36.Q;
(* Rung 43: 【Y625】B(右側) 供給ピックアップ行 *)
_e37(CLK := Out_CYw_Sply_Pick_B_F_Auto[1] AND AutoMode AND NOT Pause[1]);
_e38(CLK := Out_CYw_Sply_Pick_B_F_Manual[1] AND ManualMode);
_p39 := (_e37.Q OR _e38.Q OR Output_B_M[4]) AND NOT M9999 AND (NOT Pause[1] OR ManualMode) AND NOT Output_B_Reset_TON[4].Q;
Out_CYw_Sply_Pick_B_F := _p39;
Output_B_M[4] := _p39;
(* Rung 44 *)
Out_CYw_Sply_Pick_B_F_Done := Output_B_M[4] AND TimerQ_In_SenCY_Sply_Pick_B_F;
Output_B_Reset_TON[4](In := Output_B_M[4] AND TimerQ_In_SenCY_Sply_Pick_B_F, PT := T#1s);

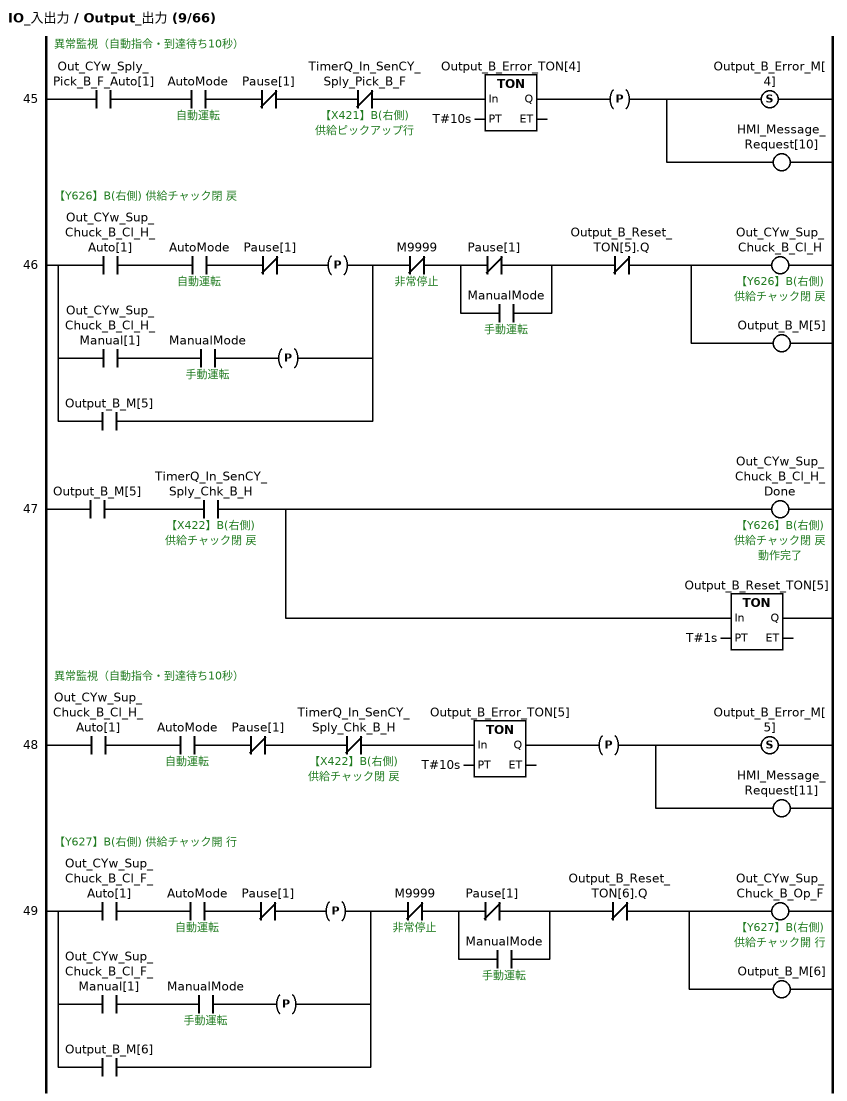
(* Rung 45: 異常監視（自動指令・到達待ち10秒） *)
Output_B_Error_TON[4](In := Out_CYw_Sply_Pick_B_F_Auto[1] AND AutoMode AND NOT Pause[1] AND NOT TimerQ_In_SenCY_Sply_Pick_B_F, PT := T#10s);
_e40(CLK := Output_B_Error_TON[4].Q);
IF _e40.Q THEN Output_B_Error_M[4] := TRUE; END_IF;
HMI_Message_Request[10] := _e40.Q;
(* Rung 46: 【Y626】B(右側) 供給チャック閉 戻 *)
_e41(CLK := Out_CYw_Sup_Chuck_B_Cl_H_Auto[1] AND AutoMode AND NOT Pause[1]);
_e42(CLK := Out_CYw_Sup_Chuck_B_Cl_H_Manual[1] AND ManualMode);
_p43 := (_e41.Q OR _e42.Q OR Output_B_M[5]) AND NOT M9999 AND (NOT Pause[1] OR ManualMode) AND NOT Output_B_Reset_TON[5].Q;
Out_CYw_Sup_Chuck_B_Cl_H := _p43;
Output_B_M[5] := _p43;
(* Rung 47 *)
Out_CYw_Sup_Chuck_B_Cl_H_Done := Output_B_M[5] AND TimerQ_In_SenCY_Sply_Chk_B_H;
Output_B_Reset_TON[5](In := Output_B_M[5] AND TimerQ_In_SenCY_Sply_Chk_B_H, PT := T#1s);
(* Rung 48: 異常監視（自動指令・到達待ち10秒） *)
Output_B_Error_TON[5](In := Out_CYw_Sup_Chuck_B_Cl_H_Auto[1] AND AutoMode AND NOT Pause[1] AND NOT TimerQ_In_SenCY_Sply_Chk_B_H, PT := T#10s);
_e44(CLK := Output_B_Error_TON[5].Q);
IF _e44.Q THEN Output_B_Error_M[5] := TRUE; END_IF;
HMI_Message_Request[11] := _e44.Q;
(* Rung 49: 【Y627】B(右側) 供給チャック開 行 *)
_e45(CLK := Out_CYw_Sup_Chuck_B_Cl_F_Auto[1] AND AutoMode AND NOT Pause[1]);
_e46(CLK := Out_CYw_Sup_Chuck_B_Cl_F_Manual[1] AND ManualMode);
_p47 := (_e45.Q OR _e46.Q OR Output_B_M[6]) AND NOT M9999 AND (NOT Pause[1] OR ManualMode) AND NOT Output_B_Reset_TON[6].Q;
Out_CYw_Sup_Chuck_B_Op_F := _p47;
Output_B_M[6] := _p47;

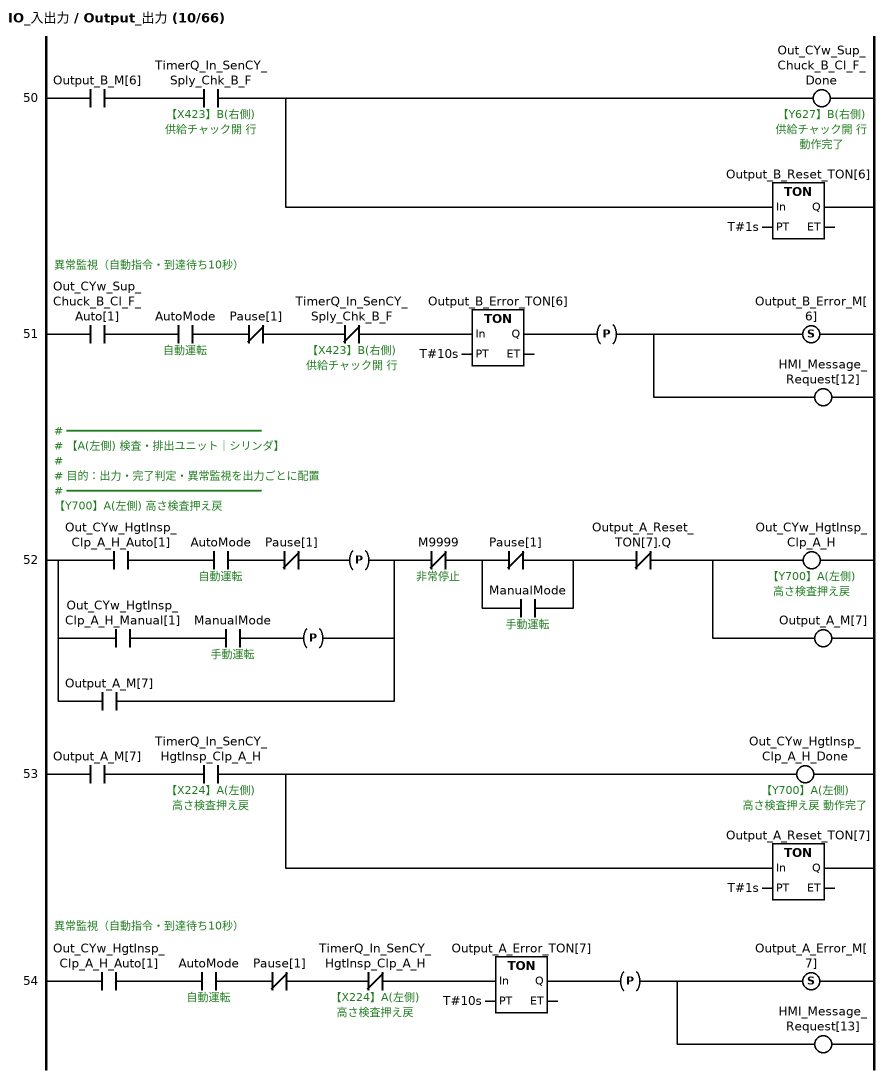
(* Rung 50 *)
Out_CYw_Sup_Chuck_B_Cl_F_Done := Output_B_M[6] AND TimerQ_In_SenCY_Sply_Chk_B_F;
Output_B_Reset_TON[6](In := Output_B_M[6] AND TimerQ_In_SenCY_Sply_Chk_B_F, PT := T#1s);
(* Rung 51: 異常監視（自動指令・到達待ち10秒） *)
Output_B_Error_TON[6](In := Out_CYw_Sup_Chuck_B_Cl_F_Auto[1] AND AutoMode AND NOT Pause[1] AND NOT TimerQ_In_SenCY_Sply_Chk_B_F, PT := T#10s);
_e48(CLK := Output_B_Error_TON[6].Q);
IF _e48.Q THEN Output_B_Error_M[6] := TRUE; END_IF;
HMI_Message_Request[12] := _e48.Q;
(* Rung 52: # ━━━━━━━━━━━━━━━━━━━━━━━━━━━━━━ / # 【A(左側) 検査・排出ユニット｜シリンダ】 / # / # 目的：出力・完了判定・異常監視を出力ごとに配置 / # ━━━━━━━━━━━━━━━━━━━━━━━━━━━━━━ / 【Y700】A(左側) 高さ検査押え戻 *)
_e49(CLK := Out_CYw_HgtInsp_Clp_A_H_Auto[1] AND AutoMode AND NOT Pause[1]);
_e50(CLK := Out_CYw_HgtInsp_Clp_A_H_Manual[1] AND ManualMode);
_p51 := (_e49.Q OR _e50.Q OR Output_A_M[7]) AND NOT M9999 AND (NOT Pause[1] OR ManualMode) AND NOT Output_A_Reset_TON[7].Q;
Out_CYw_HgtInsp_Clp_A_H := _p51;
Output_A_M[7] := _p51;
(* Rung 53 *)
_p52 := Output_A_M[7] AND TimerQ_In_SenCY_HgtInsp_Clp_A_H;
Out_CYw_HgtInsp_Clp_A_H_Done := _p52;
Output_A_Reset_TON[7](In := _p52, PT := T#1s);
(* Rung 54: 異常監視（自動指令・到達待ち10秒） *)
Output_A_Error_TON[7](In := Out_CYw_HgtInsp_Clp_A_H_Auto[1] AND AutoMode AND NOT Pause[1] AND NOT TimerQ_In_SenCY_HgtInsp_Clp_A_H, PT := T#10s);
_e53(CLK := Output_A_Error_TON[7].Q);
IF _e53.Q THEN Output_A_Error_M[7] := TRUE; END_IF;
HMI_Message_Request[13] := _e53.Q;

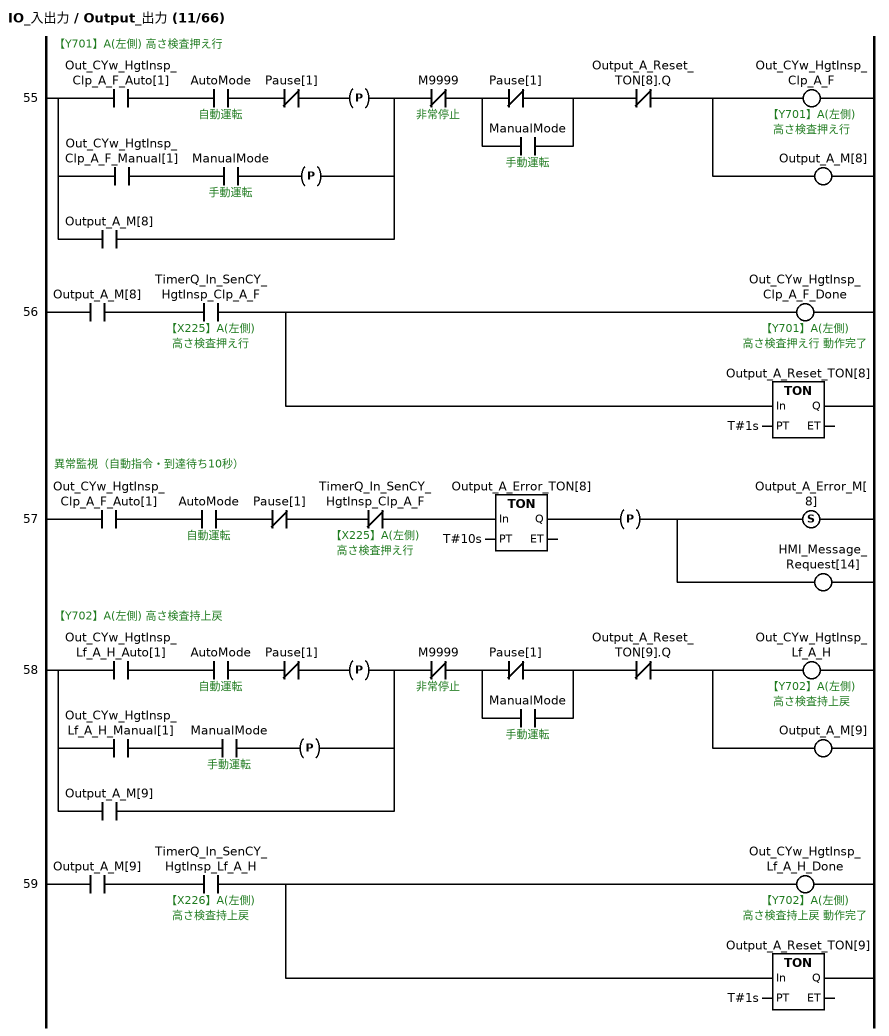
(* Rung 55: 【Y701】A(左側) 高さ検査押え行 *)
_e54(CLK := Out_CYw_HgtInsp_Clp_A_F_Auto[1] AND AutoMode AND NOT Pause[1]);
_e55(CLK := Out_CYw_HgtInsp_Clp_A_F_Manual[1] AND ManualMode);
_p56 := (_e54.Q OR _e55.Q OR Output_A_M[8]) AND NOT M9999 AND (NOT Pause[1] OR ManualMode) AND NOT Output_A_Reset_TON[8].Q;
Out_CYw_HgtInsp_Clp_A_F := _p56;
Output_A_M[8] := _p56;
(* Rung 56 *)
_p57 := Output_A_M[8] AND TimerQ_In_SenCY_HgtInsp_Clp_A_F;
Out_CYw_HgtInsp_Clp_A_F_Done := _p57;
Output_A_Reset_TON[8](In := _p57, PT := T#1s);
(* Rung 57: 異常監視（自動指令・到達待ち10秒） *)
Output_A_Error_TON[8](In := Out_CYw_HgtInsp_Clp_A_F_Auto[1] AND AutoMode AND NOT Pause[1] AND NOT TimerQ_In_SenCY_HgtInsp_Clp_A_F, PT := T#10s);
_e58(CLK := Output_A_Error_TON[8].Q);
IF _e58.Q THEN Output_A_Error_M[8] := TRUE; END_IF;
HMI_Message_Request[14] := _e58.Q;
(* Rung 58: 【Y702】A(左側) 高さ検査持上戻 *)
_e59(CLK := Out_CYw_HgtInsp_Lf_A_H_Auto[1] AND AutoMode AND NOT Pause[1]);
_e60(CLK := Out_CYw_HgtInsp_Lf_A_H_Manual[1] AND ManualMode);
_p61 := (_e59.Q OR _e60.Q OR Output_A_M[9]) AND NOT M9999 AND (NOT Pause[1] OR ManualMode) AND NOT Output_A_Reset_TON[9].Q;
Out_CYw_HgtInsp_Lf_A_H := _p61;
Output_A_M[9] := _p61;
(* Rung 59 *)
Out_CYw_HgtInsp_Lf_A_H_Done := Output_A_M[9] AND TimerQ_In_SenCY_HgtInsp_Lf_A_H;
Output_A_Reset_TON[9](In := Output_A_M[9] AND TimerQ_In_SenCY_HgtInsp_Lf_A_H, PT := T#1s);

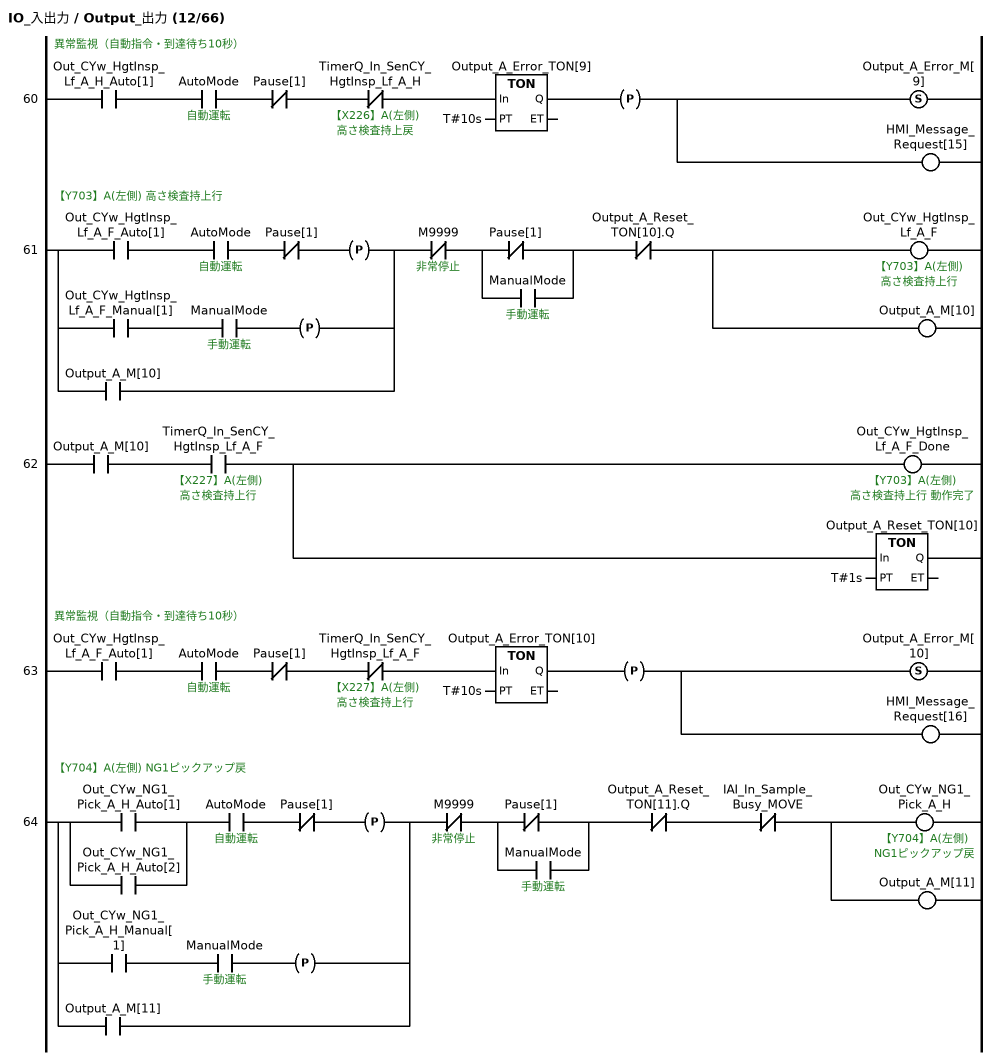
(* Rung 60: 異常監視（自動指令・到達待ち10秒） *)
Output_A_Error_TON[9](In := Out_CYw_HgtInsp_Lf_A_H_Auto[1] AND AutoMode AND NOT Pause[1] AND NOT TimerQ_In_SenCY_HgtInsp_Lf_A_H, PT := T#10s);
_e62(CLK := Output_A_Error_TON[9].Q);
IF _e62.Q THEN Output_A_Error_M[9] := TRUE; END_IF;
HMI_Message_Request[15] := _e62.Q;
(* Rung 61: 【Y703】A(左側) 高さ検査持上行 *)
_e63(CLK := Out_CYw_HgtInsp_Lf_A_F_Auto[1] AND AutoMode AND NOT Pause[1]);
_e64(CLK := Out_CYw_HgtInsp_Lf_A_F_Manual[1] AND ManualMode);
_p65 := (_e63.Q OR _e64.Q OR Output_A_M[10]) AND NOT M9999 AND (NOT Pause[1] OR ManualMode) AND NOT Output_A_Reset_TON[10].Q;
Out_CYw_HgtInsp_Lf_A_F := _p65;
Output_A_M[10] := _p65;
(* Rung 62 *)
_p66 := Output_A_M[10] AND TimerQ_In_SenCY_HgtInsp_Lf_A_F;
Out_CYw_HgtInsp_Lf_A_F_Done := _p66;
Output_A_Reset_TON[10](In := _p66, PT := T#1s);
(* Rung 63: 異常監視（自動指令・到達待ち10秒） *)
Output_A_Error_TON[10](In := Out_CYw_HgtInsp_Lf_A_F_Auto[1] AND AutoMode AND NOT Pause[1] AND NOT TimerQ_In_SenCY_HgtInsp_Lf_A_F, PT := T#10s);
_e67(CLK := Output_A_Error_TON[10].Q);
IF _e67.Q THEN Output_A_Error_M[10] := TRUE; END_IF;
HMI_Message_Request[16] := _e67.Q;
(* Rung 64: 【Y704】A(左側) NG1ピックアップ戻 *)
_e68(CLK := (Out_CYw_NG1_Pick_A_H_Auto[1] OR Out_CYw_NG1_Pick_A_H_Auto[2]) AND AutoMode AND NOT Pause[1]);
_e69(CLK := Out_CYw_NG1_Pick_A_H_Manual[1] AND ManualMode);
_p70 := (_e68.Q OR _e69.Q OR Output_A_M[11]) AND NOT M9999 AND (NOT Pause[1] OR ManualMode) AND NOT Output_A_Reset_TON[11].Q AND NOT IAI_In_Sample_Busy_MOVE;
Out_CYw_NG1_Pick_A_H := _p70;
Output_A_M[11] := _p70;

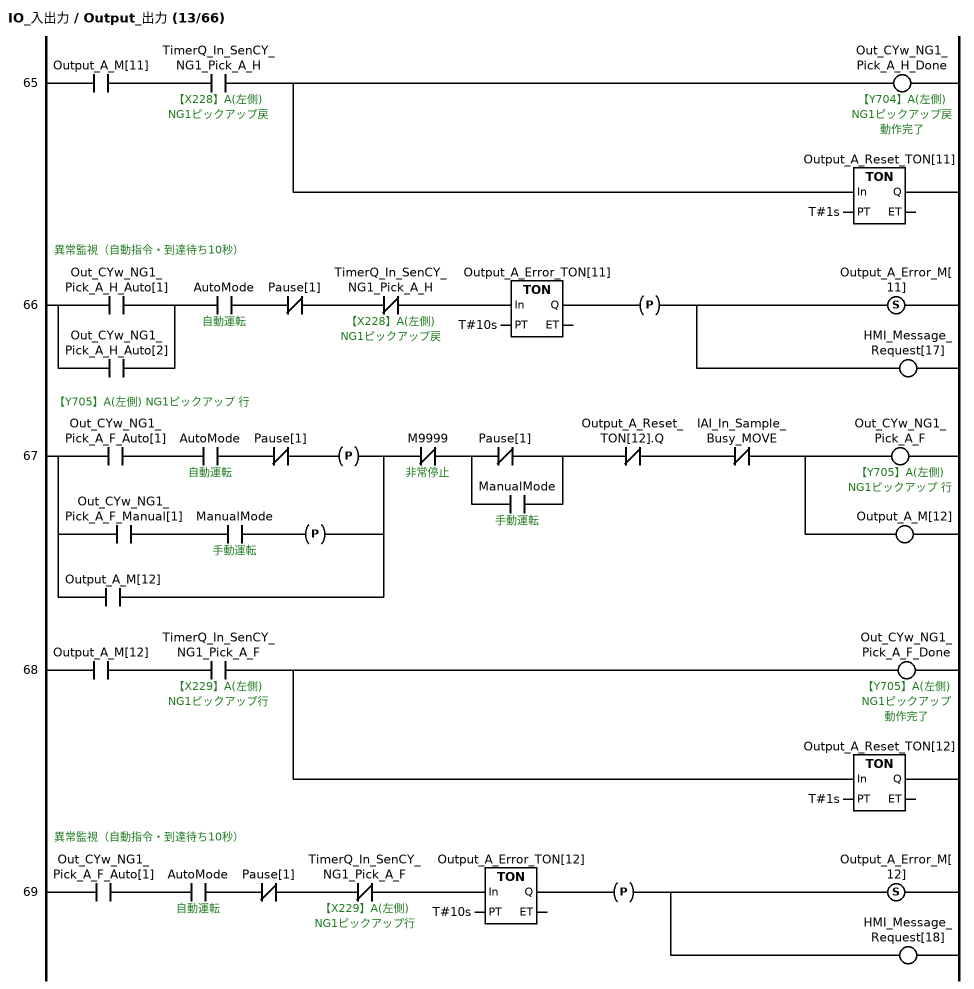
(* Rung 65 *)
Out_CYw_NG1_Pick_A_H_Done := Output_A_M[11] AND TimerQ_In_SenCY_NG1_Pick_A_H;
Output_A_Reset_TON[11](In := Output_A_M[11] AND TimerQ_In_SenCY_NG1_Pick_A_H, PT := T#1s);
(* Rung 66: 異常監視（自動指令・到達待ち10秒） *)
Output_A_Error_TON[11](In := (Out_CYw_NG1_Pick_A_H_Auto[1] OR Out_CYw_NG1_Pick_A_H_Auto[2]) AND AutoMode AND NOT Pause[1] AND NOT TimerQ_In_SenCY_NG1_Pick_A_H, PT := T#10s);
_e71(CLK := Output_A_Error_TON[11].Q);
IF _e71.Q THEN Output_A_Error_M[11] := TRUE; END_IF;
HMI_Message_Request[17] := _e71.Q;
(* Rung 67: 【Y705】A(左側) NG1ピックアップ 行 *)
_e72(CLK := Out_CYw_NG1_Pick_A_F_Auto[1] AND AutoMode AND NOT Pause[1]);
_e73(CLK := Out_CYw_NG1_Pick_A_F_Manual[1] AND ManualMode);
_p74 := (_e72.Q OR _e73.Q OR Output_A_M[12]) AND NOT M9999 AND (NOT Pause[1] OR ManualMode) AND NOT Output_A_Reset_TON[12].Q AND NOT IAI_In_Sample_Busy_MOVE;
Out_CYw_NG1_Pick_A_F := _p74;
Output_A_M[12] := _p74;
(* Rung 68 *)
Out_CYw_NG1_Pick_A_F_Done := Output_A_M[12] AND TimerQ_In_SenCY_NG1_Pick_A_F;
Output_A_Reset_TON[12](In := Output_A_M[12] AND TimerQ_In_SenCY_NG1_Pick_A_F, PT := T#1s);
(* Rung 69: 異常監視（自動指令・到達待ち10秒） *)
Output_A_Error_TON[12](In := Out_CYw_NG1_Pick_A_F_Auto[1] AND AutoMode AND NOT Pause[1] AND NOT TimerQ_In_SenCY_NG1_Pick_A_F, PT := T#10s);
_e75(CLK := Output_A_Error_TON[12].Q);
IF _e75.Q THEN Output_A_Error_M[12] := TRUE; END_IF;
HMI_Message_Request[18] := _e75.Q;

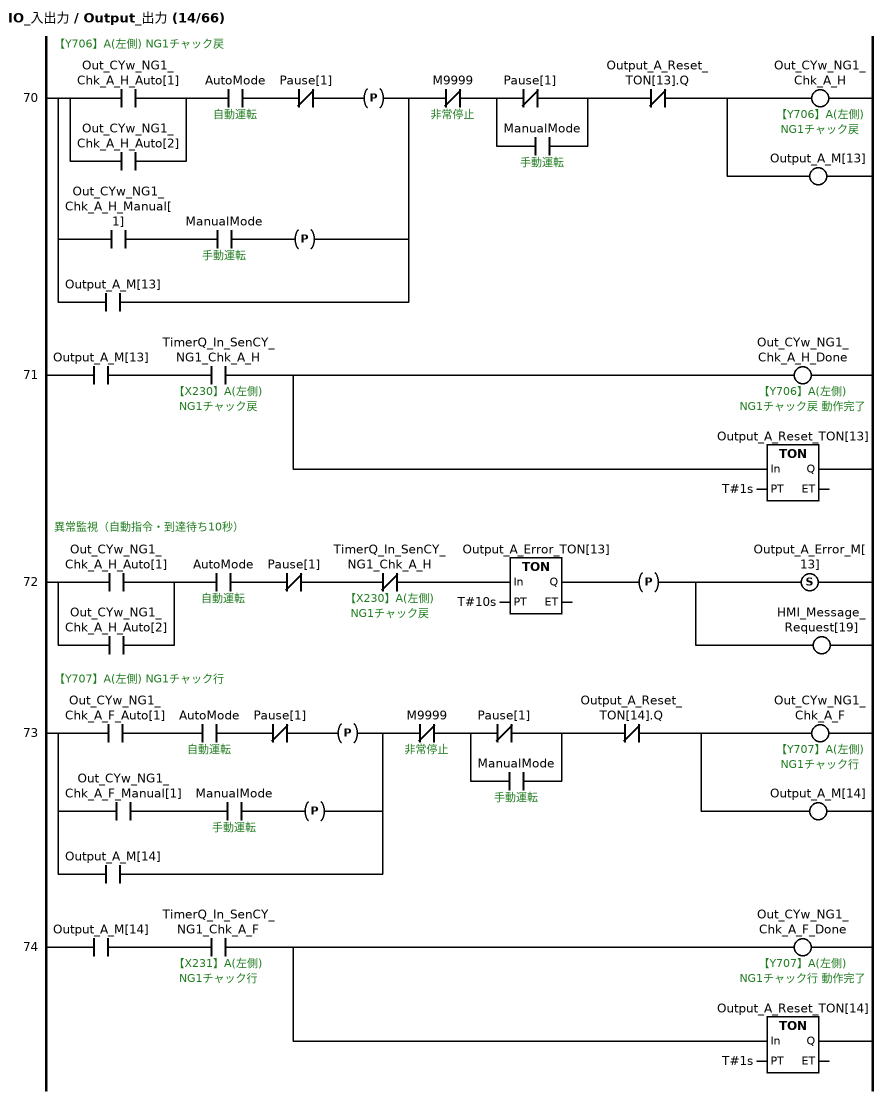
(* Rung 70: 【Y706】A(左側) NG1チャック戻 *)
_e76(CLK := (Out_CYw_NG1_Chk_A_H_Auto[1] OR Out_CYw_NG1_Chk_A_H_Auto[2]) AND AutoMode AND NOT Pause[1]);
_e77(CLK := Out_CYw_NG1_Chk_A_H_Manual[1] AND ManualMode);
_p78 := (_e76.Q OR _e77.Q OR Output_A_M[13]) AND NOT M9999 AND (NOT Pause[1] OR ManualMode) AND NOT Output_A_Reset_TON[13].Q;
Out_CYw_NG1_Chk_A_H := _p78;
Output_A_M[13] := _p78;
(* Rung 71 *)
Out_CYw_NG1_Chk_A_H_Done := Output_A_M[13] AND TimerQ_In_SenCY_NG1_Chk_A_H;
Output_A_Reset_TON[13](In := Output_A_M[13] AND TimerQ_In_SenCY_NG1_Chk_A_H, PT := T#1s);
(* Rung 72: 異常監視（自動指令・到達待ち10秒） *)
Output_A_Error_TON[13](In := (Out_CYw_NG1_Chk_A_H_Auto[1] OR Out_CYw_NG1_Chk_A_H_Auto[2]) AND AutoMode AND NOT Pause[1] AND NOT TimerQ_In_SenCY_NG1_Chk_A_H, PT := T#10s);
_e79(CLK := Output_A_Error_TON[13].Q);
IF _e79.Q THEN Output_A_Error_M[13] := TRUE; END_IF;
HMI_Message_Request[19] := _e79.Q;
(* Rung 73: 【Y707】A(左側) NG1チャック行 *)
_e80(CLK := Out_CYw_NG1_Chk_A_F_Auto[1] AND AutoMode AND NOT Pause[1]);
_e81(CLK := Out_CYw_NG1_Chk_A_F_Manual[1] AND ManualMode);
_p82 := (_e80.Q OR _e81.Q OR Output_A_M[14]) AND NOT M9999 AND (NOT Pause[1] OR ManualMode) AND NOT Output_A_Reset_TON[14].Q;
Out_CYw_NG1_Chk_A_F := _p82;
Output_A_M[14] := _p82;
(* Rung 74 *)
Out_CYw_NG1_Chk_A_F_Done := Output_A_M[14] AND TimerQ_In_SenCY_NG1_Chk_A_F;
Output_A_Reset_TON[14](In := Output_A_M[14] AND TimerQ_In_SenCY_NG1_Chk_A_F, PT := T#1s);

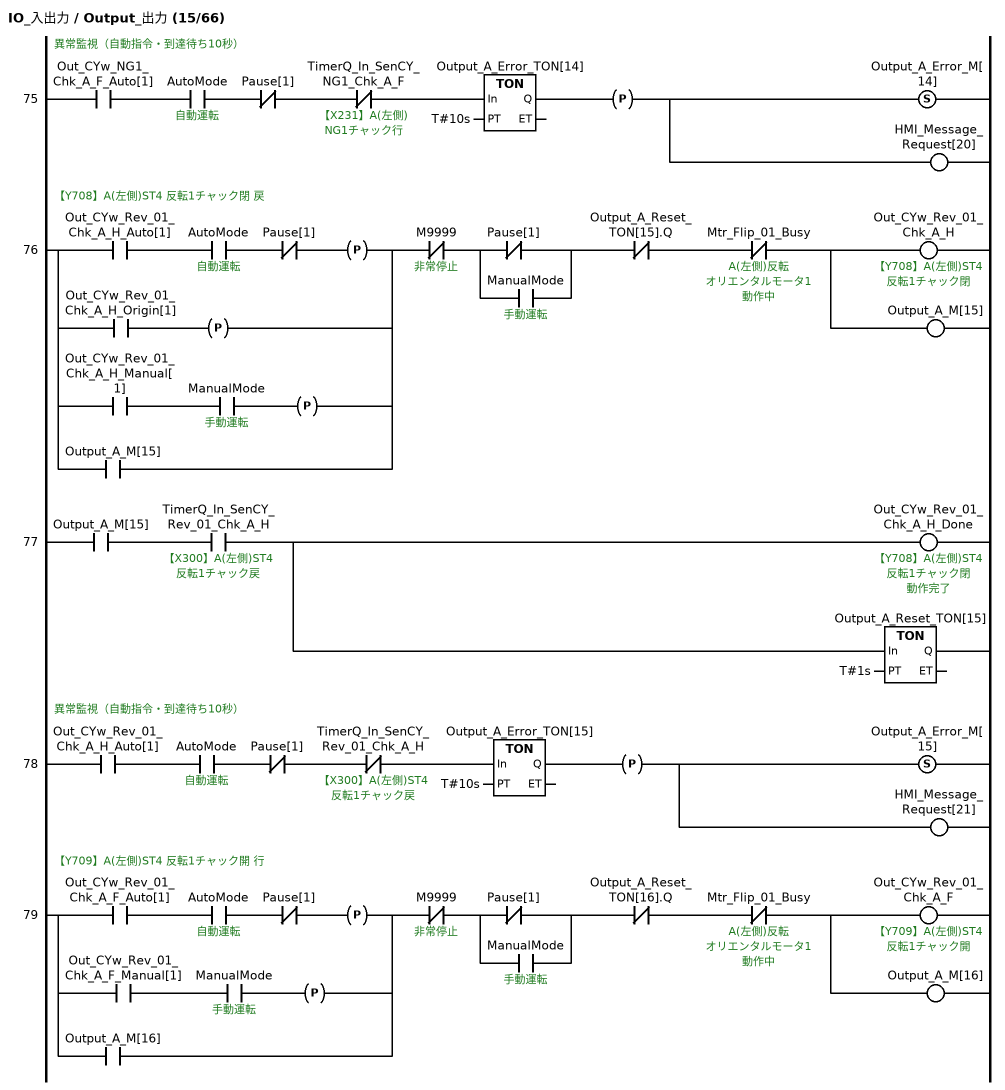
(* Rung 75: 異常監視（自動指令・到達待ち10秒） *)
Output_A_Error_TON[14](In := Out_CYw_NG1_Chk_A_F_Auto[1] AND AutoMode AND NOT Pause[1] AND NOT TimerQ_In_SenCY_NG1_Chk_A_F, PT := T#10s);
_e83(CLK := Output_A_Error_TON[14].Q);
IF _e83.Q THEN Output_A_Error_M[14] := TRUE; END_IF;
HMI_Message_Request[20] := _e83.Q;
(* Rung 76: 【Y708】A(左側)ST4 反転1チャック閉 戻 *)
_e84(CLK := Out_CYw_Rev_01_Chk_A_H_Auto[1] AND AutoMode AND NOT Pause[1]);
_e85(CLK := Out_CYw_Rev_01_Chk_A_H_Origin[1]);
_e86(CLK := Out_CYw_Rev_01_Chk_A_H_Manual[1] AND ManualMode);
_p87 := (_e84.Q OR _e85.Q OR _e86.Q OR Output_A_M[15]) AND NOT M9999 AND (NOT Pause[1] OR ManualMode) AND NOT Output_A_Reset_TON[15].Q AND NOT Mtr_Flip_01_Busy;
Out_CYw_Rev_01_Chk_A_H := _p87;
Output_A_M[15] := _p87;
(* Rung 77 *)
_p88 := Output_A_M[15] AND TimerQ_In_SenCY_Rev_01_Chk_A_H;
Out_CYw_Rev_01_Chk_A_H_Done := _p88;
Output_A_Reset_TON[15](In := _p88, PT := T#1s);
(* Rung 78: 異常監視（自動指令・到達待ち10秒） *)
Output_A_Error_TON[15](In := Out_CYw_Rev_01_Chk_A_H_Auto[1] AND AutoMode AND NOT Pause[1] AND NOT TimerQ_In_SenCY_Rev_01_Chk_A_H, PT := T#10s);
_e89(CLK := Output_A_Error_TON[15].Q);
IF _e89.Q THEN Output_A_Error_M[15] := TRUE; END_IF;
HMI_Message_Request[21] := _e89.Q;
(* Rung 79: 【Y709】A(左側)ST4 反転1チャック開 行 *)
_e90(CLK := Out_CYw_Rev_01_Chk_A_F_Auto[1] AND AutoMode AND NOT Pause[1]);
_e91(CLK := Out_CYw_Rev_01_Chk_A_F_Manual[1] AND ManualMode);
_p92 := (_e90.Q OR _e91.Q OR Output_A_M[16]) AND NOT M9999 AND (NOT Pause[1] OR ManualMode) AND NOT Output_A_Reset_TON[16].Q AND NOT Mtr_Flip_01_Busy;
Out_CYw_Rev_01_Chk_A_F := _p92;
Output_A_M[16] := _p92;

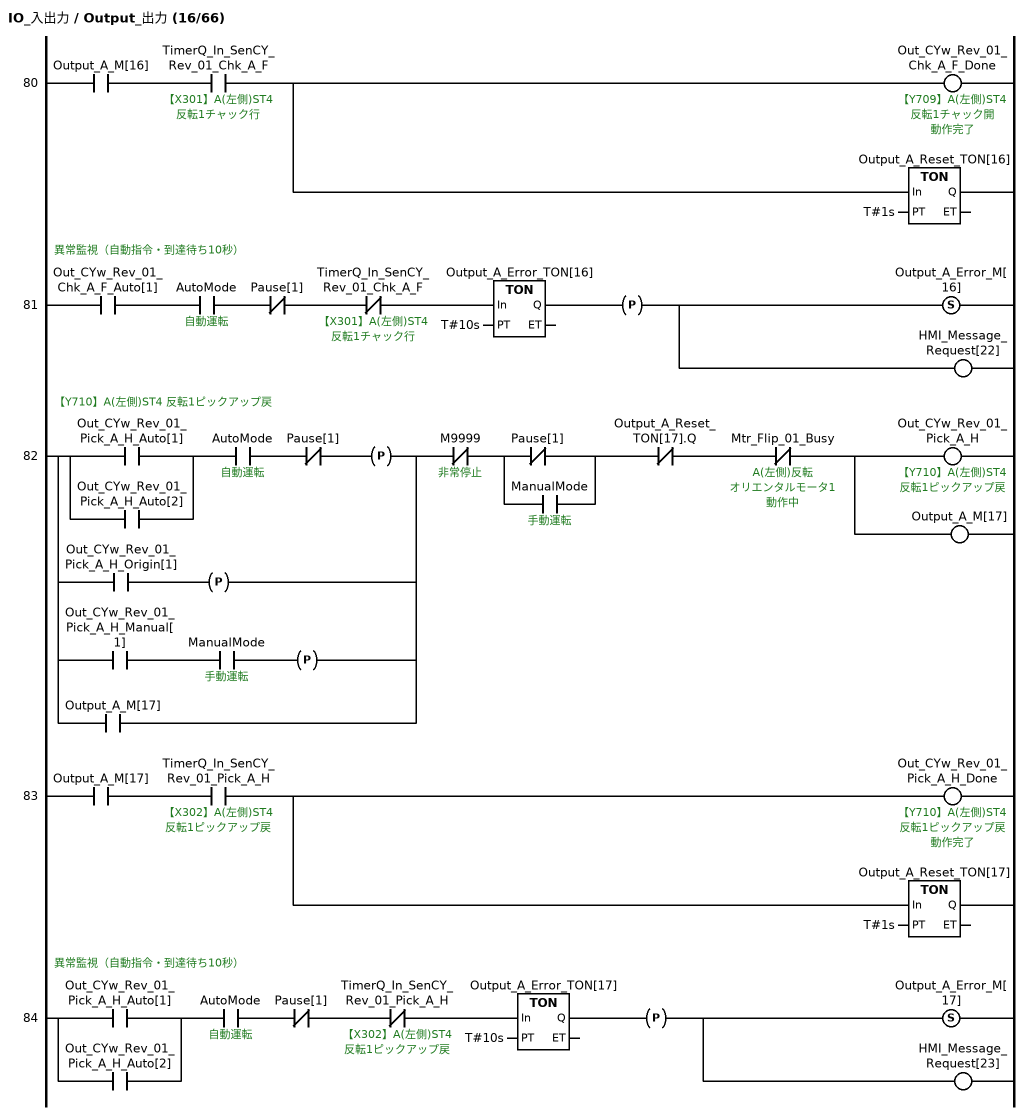
(* Rung 80 *)
_p93 := Output_A_M[16] AND TimerQ_In_SenCY_Rev_01_Chk_A_F;
Out_CYw_Rev_01_Chk_A_F_Done := _p93;
Output_A_Reset_TON[16](In := _p93, PT := T#1s);
(* Rung 81: 異常監視（自動指令・到達待ち10秒） *)
Output_A_Error_TON[16](In := Out_CYw_Rev_01_Chk_A_F_Auto[1] AND AutoMode AND NOT Pause[1] AND NOT TimerQ_In_SenCY_Rev_01_Chk_A_F, PT := T#10s);
_e94(CLK := Output_A_Error_TON[16].Q);
IF _e94.Q THEN Output_A_Error_M[16] := TRUE; END_IF;
HMI_Message_Request[22] := _e94.Q;
(* Rung 82: 【Y710】A(左側)ST4 反転1ピックアップ戻 *)
_e95(CLK := (Out_CYw_Rev_01_Pick_A_H_Auto[1] OR Out_CYw_Rev_01_Pick_A_H_Auto[2]) AND AutoMode AND NOT Pause[1]);
_e96(CLK := Out_CYw_Rev_01_Pick_A_H_Origin[1]);
_e97(CLK := Out_CYw_Rev_01_Pick_A_H_Manual[1] AND ManualMode);
_p98 := (_e95.Q OR _e96.Q OR _e97.Q OR Output_A_M[17]) AND NOT M9999 AND (NOT Pause[1] OR ManualMode) AND NOT Output_A_Reset_TON[17].Q AND NOT Mtr_Flip_01_Busy;
Out_CYw_Rev_01_Pick_A_H := _p98;
Output_A_M[17] := _p98;
(* Rung 83 *)
_p99 := Output_A_M[17] AND TimerQ_In_SenCY_Rev_01_Pick_A_H;
Out_CYw_Rev_01_Pick_A_H_Done := _p99;
Output_A_Reset_TON[17](In := _p99, PT := T#1s);
(* Rung 84: 異常監視（自動指令・到達待ち10秒） *)
Output_A_Error_TON[17](In := (Out_CYw_Rev_01_Pick_A_H_Auto[1] OR Out_CYw_Rev_01_Pick_A_H_Auto[2]) AND AutoMode AND NOT Pause[1] AND NOT TimerQ_In_SenCY_Rev_01_Pick_A_H, PT := T#10s);
_e100(CLK := Output_A_Error_TON[17].Q);
IF _e100.Q THEN Output_A_Error_M[17] := TRUE; END_IF;
HMI_Message_Request[23] := _e100.Q;

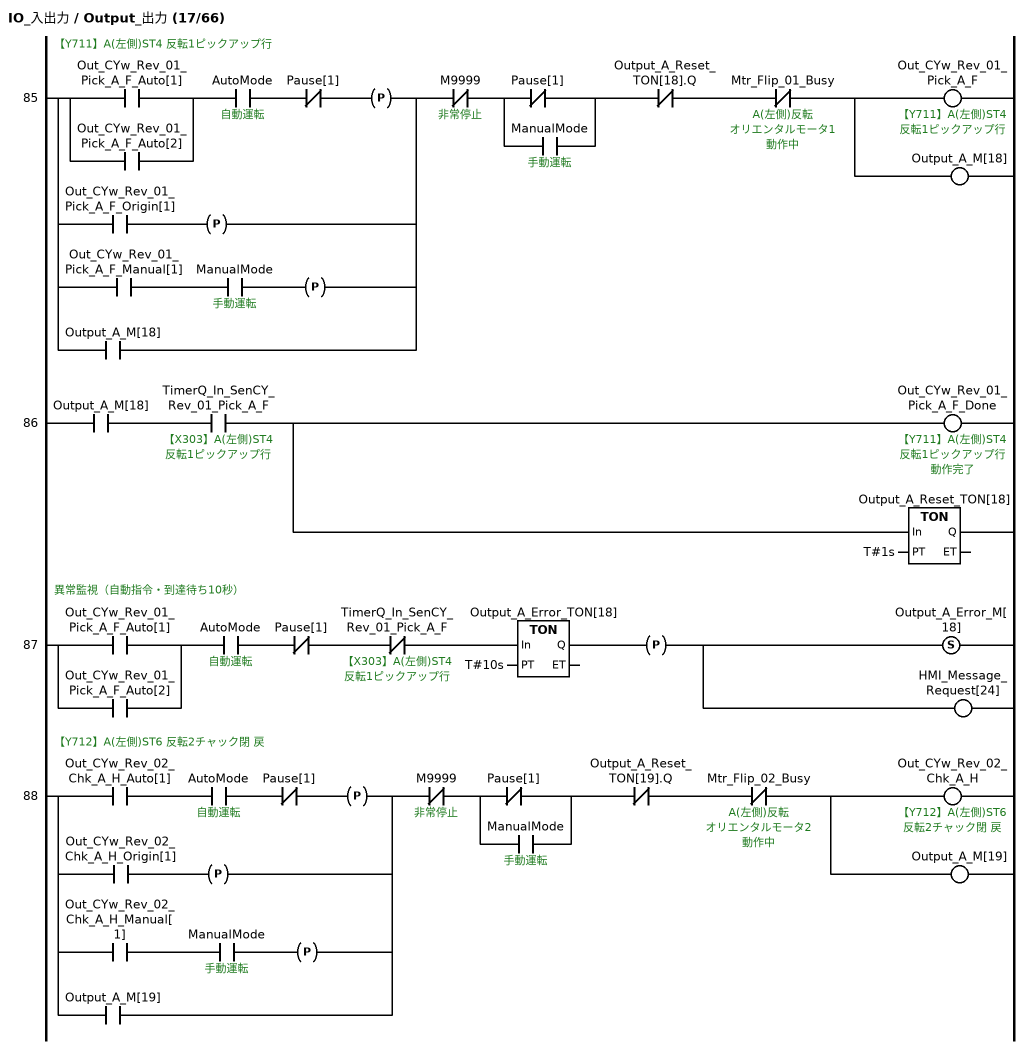
(* Rung 85: 【Y711】A(左側)ST4 反転1ピックアップ行 *)
_e101(CLK := (Out_CYw_Rev_01_Pick_A_F_Auto[1] OR Out_CYw_Rev_01_Pick_A_F_Auto[2]) AND AutoMode AND NOT Pause[1]);
_e102(CLK := Out_CYw_Rev_01_Pick_A_F_Origin[1]);
_e103(CLK := Out_CYw_Rev_01_Pick_A_F_Manual[1] AND ManualMode);
_p104 := (_e101.Q OR _e102.Q OR _e103.Q OR Output_A_M[18]) AND NOT M9999 AND (NOT Pause[1] OR ManualMode) AND NOT Output_A_Reset_TON[18].Q AND NOT Mtr_Flip_01_Busy;
Out_CYw_Rev_01_Pick_A_F := _p104;
Output_A_M[18] := _p104;
(* Rung 86 *)
_p105 := Output_A_M[18] AND TimerQ_In_SenCY_Rev_01_Pick_A_F;
Out_CYw_Rev_01_Pick_A_F_Done := _p105;
Output_A_Reset_TON[18](In := _p105, PT := T#1s);
(* Rung 87: 異常監視（自動指令・到達待ち10秒） *)
Output_A_Error_TON[18](In := (Out_CYw_Rev_01_Pick_A_F_Auto[1] OR Out_CYw_Rev_01_Pick_A_F_Auto[2]) AND AutoMode AND NOT Pause[1] AND NOT TimerQ_In_SenCY_Rev_01_Pick_A_F, PT := T#10s);
_e106(CLK := Output_A_Error_TON[18].Q);
IF _e106.Q THEN Output_A_Error_M[18] := TRUE; END_IF;
HMI_Message_Request[24] := _e106.Q;
(* Rung 88: 【Y712】A(左側)ST6 反転2チャック閉 戻 *)
_e107(CLK := Out_CYw_Rev_02_Chk_A_H_Auto[1] AND AutoMode AND NOT Pause[1]);
_e108(CLK := Out_CYw_Rev_02_Chk_A_H_Origin[1]);
_e109(CLK := Out_CYw_Rev_02_Chk_A_H_Manual[1] AND ManualMode);
_p110 := (_e107.Q OR _e108.Q OR _e109.Q OR Output_A_M[19]) AND NOT M9999 AND (NOT Pause[1] OR ManualMode) AND NOT Output_A_Reset_TON[19].Q AND NOT Mtr_Flip_02_Busy;
Out_CYw_Rev_02_Chk_A_H := _p110;
Output_A_M[19] := _p110;

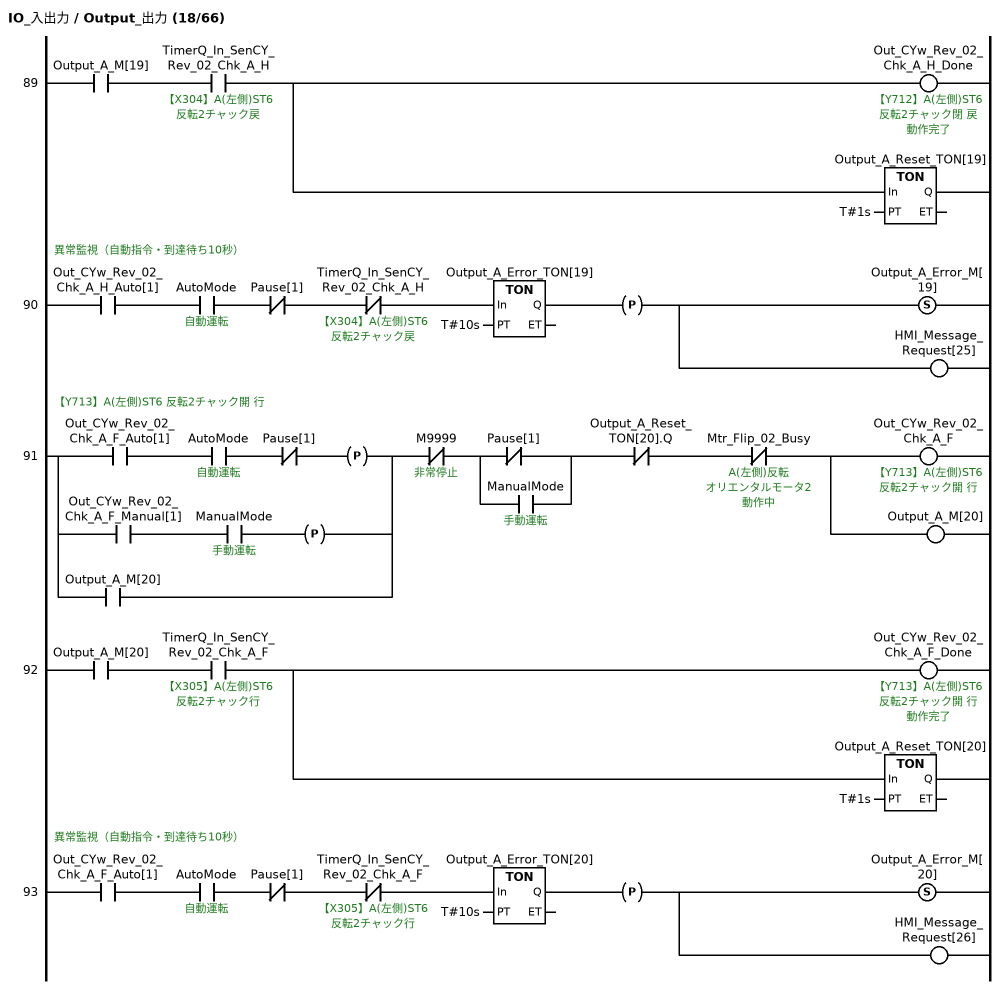
(* Rung 89 *)
_p111 := Output_A_M[19] AND TimerQ_In_SenCY_Rev_02_Chk_A_H;
Out_CYw_Rev_02_Chk_A_H_Done := _p111;
Output_A_Reset_TON[19](In := _p111, PT := T#1s);
(* Rung 90: 異常監視（自動指令・到達待ち10秒） *)
Output_A_Error_TON[19](In := Out_CYw_Rev_02_Chk_A_H_Auto[1] AND AutoMode AND NOT Pause[1] AND NOT TimerQ_In_SenCY_Rev_02_Chk_A_H, PT := T#10s);
_e112(CLK := Output_A_Error_TON[19].Q);
IF _e112.Q THEN Output_A_Error_M[19] := TRUE; END_IF;
HMI_Message_Request[25] := _e112.Q;
(* Rung 91: 【Y713】A(左側)ST6 反転2チャック開 行 *)
_e113(CLK := Out_CYw_Rev_02_Chk_A_F_Auto[1] AND AutoMode AND NOT Pause[1]);
_e114(CLK := Out_CYw_Rev_02_Chk_A_F_Manual[1] AND ManualMode);
_p115 := (_e113.Q OR _e114.Q OR Output_A_M[20]) AND NOT M9999 AND (NOT Pause[1] OR ManualMode) AND NOT Output_A_Reset_TON[20].Q AND NOT Mtr_Flip_02_Busy;
Out_CYw_Rev_02_Chk_A_F := _p115;
Output_A_M[20] := _p115;
(* Rung 92 *)
_p116 := Output_A_M[20] AND TimerQ_In_SenCY_Rev_02_Chk_A_F;
Out_CYw_Rev_02_Chk_A_F_Done := _p116;
Output_A_Reset_TON[20](In := _p116, PT := T#1s);
(* Rung 93: 異常監視（自動指令・到達待ち10秒） *)
Output_A_Error_TON[20](In := Out_CYw_Rev_02_Chk_A_F_Auto[1] AND AutoMode AND NOT Pause[1] AND NOT TimerQ_In_SenCY_Rev_02_Chk_A_F, PT := T#10s);
_e117(CLK := Output_A_Error_TON[20].Q);
IF _e117.Q THEN Output_A_Error_M[20] := TRUE; END_IF;
HMI_Message_Request[26] := _e117.Q;

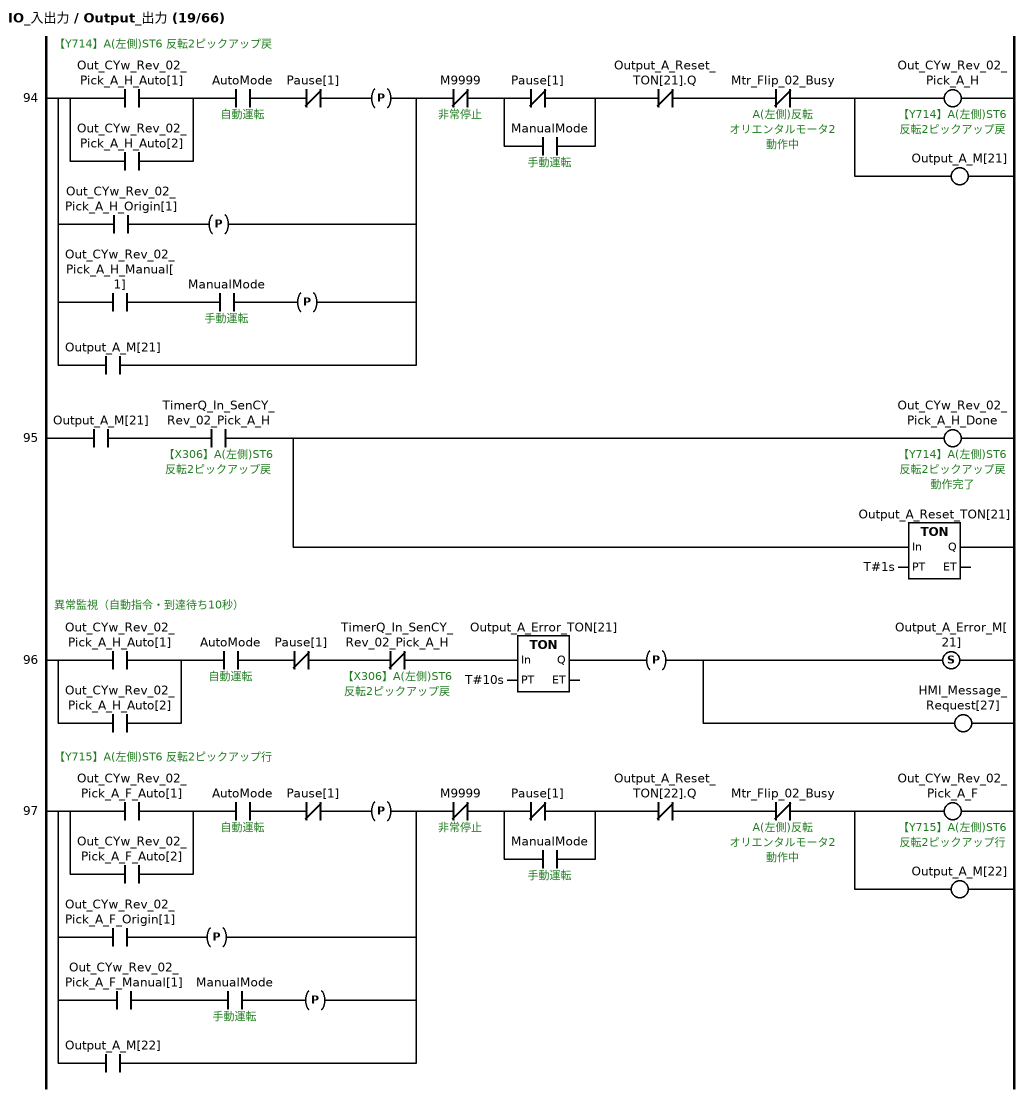
(* Rung 94: 【Y714】A(左側)ST6 反転2ピックアップ戻 *)
_e118(CLK := (Out_CYw_Rev_02_Pick_A_H_Auto[1] OR Out_CYw_Rev_02_Pick_A_H_Auto[2]) AND AutoMode AND NOT Pause[1]);
_e119(CLK := Out_CYw_Rev_02_Pick_A_H_Origin[1]);
_e120(CLK := Out_CYw_Rev_02_Pick_A_H_Manual[1] AND ManualMode);
_p121 := (_e118.Q OR _e119.Q OR _e120.Q OR Output_A_M[21]) AND NOT M9999 AND (NOT Pause[1] OR ManualMode) AND NOT Output_A_Reset_TON[21].Q AND NOT Mtr_Flip_02_Busy;
Out_CYw_Rev_02_Pick_A_H := _p121;
Output_A_M[21] := _p121;
(* Rung 95 *)
_p122 := Output_A_M[21] AND TimerQ_In_SenCY_Rev_02_Pick_A_H;
Out_CYw_Rev_02_Pick_A_H_Done := _p122;
Output_A_Reset_TON[21](In := _p122, PT := T#1s);
(* Rung 96: 異常監視（自動指令・到達待ち10秒） *)
Output_A_Error_TON[21](In := (Out_CYw_Rev_02_Pick_A_H_Auto[1] OR Out_CYw_Rev_02_Pick_A_H_Auto[2]) AND AutoMode AND NOT Pause[1] AND NOT TimerQ_In_SenCY_Rev_02_Pick_A_H, PT := T#10s);
_e123(CLK := Output_A_Error_TON[21].Q);
IF _e123.Q THEN Output_A_Error_M[21] := TRUE; END_IF;
HMI_Message_Request[27] := _e123.Q;
(* Rung 97: 【Y715】A(左側)ST6 反転2ピックアップ行 *)
_e124(CLK := (Out_CYw_Rev_02_Pick_A_F_Auto[1] OR Out_CYw_Rev_02_Pick_A_F_Auto[2]) AND AutoMode AND NOT Pause[1]);
_e125(CLK := Out_CYw_Rev_02_Pick_A_F_Origin[1]);
_e126(CLK := Out_CYw_Rev_02_Pick_A_F_Manual[1] AND ManualMode);
_p127 := (_e124.Q OR _e125.Q OR _e126.Q OR Output_A_M[22]) AND NOT M9999 AND (NOT Pause[1] OR ManualMode) AND NOT Output_A_Reset_TON[22].Q AND NOT Mtr_Flip_02_Busy;
Out_CYw_Rev_02_Pick_A_F := _p127;
Output_A_M[22] := _p127;

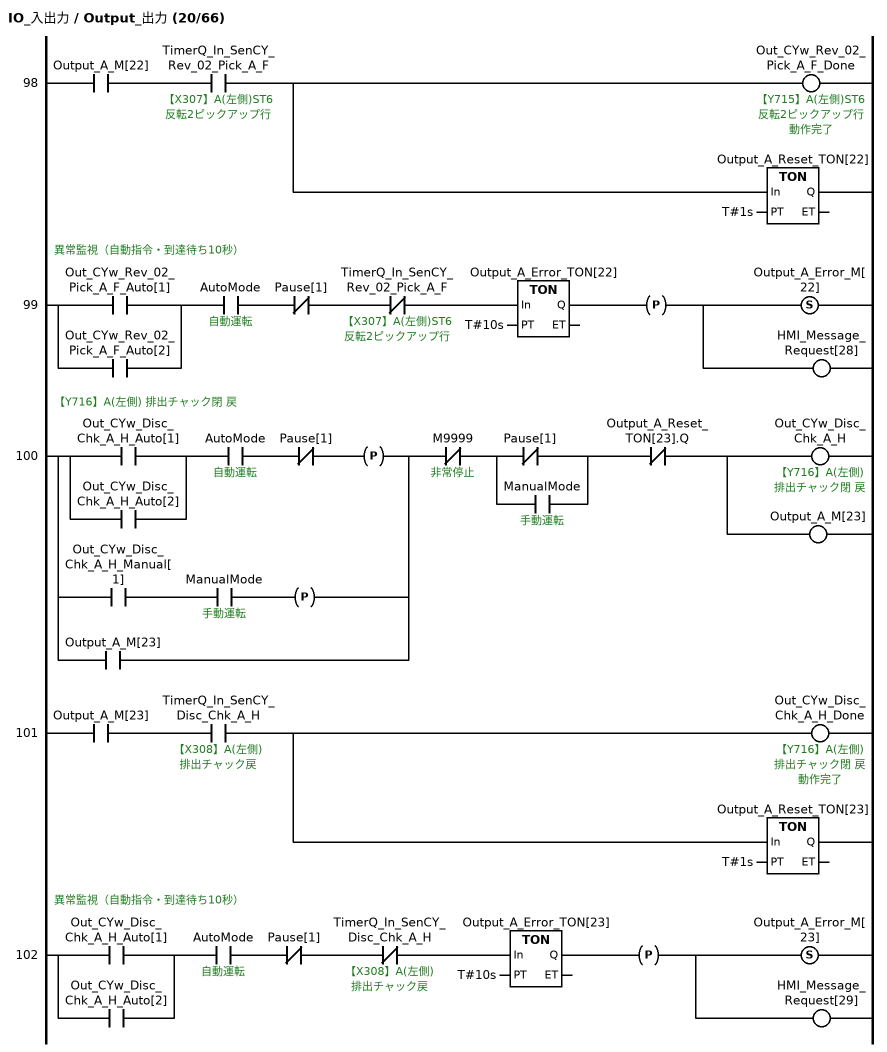
(* Rung 98 *)
_p128 := Output_A_M[22] AND TimerQ_In_SenCY_Rev_02_Pick_A_F;
Out_CYw_Rev_02_Pick_A_F_Done := _p128;
Output_A_Reset_TON[22](In := _p128, PT := T#1s);
(* Rung 99: 異常監視（自動指令・到達待ち10秒） *)
Output_A_Error_TON[22](In := (Out_CYw_Rev_02_Pick_A_F_Auto[1] OR Out_CYw_Rev_02_Pick_A_F_Auto[2]) AND AutoMode AND NOT Pause[1] AND NOT TimerQ_In_SenCY_Rev_02_Pick_A_F, PT := T#10s);
_e129(CLK := Output_A_Error_TON[22].Q);
IF _e129.Q THEN Output_A_Error_M[22] := TRUE; END_IF;
HMI_Message_Request[28] := _e129.Q;
(* Rung 100: 【Y716】A(左側) 排出チャック閉 戻 *)
_e130(CLK := (Out_CYw_Disc_Chk_A_H_Auto[1] OR Out_CYw_Disc_Chk_A_H_Auto[2]) AND AutoMode AND NOT Pause[1]);
_e131(CLK := Out_CYw_Disc_Chk_A_H_Manual[1] AND ManualMode);
_p132 := (_e130.Q OR _e131.Q OR Output_A_M[23]) AND NOT M9999 AND (NOT Pause[1] OR ManualMode) AND NOT Output_A_Reset_TON[23].Q;
Out_CYw_Disc_Chk_A_H := _p132;
Output_A_M[23] := _p132;
(* Rung 101 *)
Out_CYw_Disc_Chk_A_H_Done := Output_A_M[23] AND TimerQ_In_SenCY_Disc_Chk_A_H;
Output_A_Reset_TON[23](In := Output_A_M[23] AND TimerQ_In_SenCY_Disc_Chk_A_H, PT := T#1s);
(* Rung 102: 異常監視（自動指令・到達待ち10秒） *)
Output_A_Error_TON[23](In := (Out_CYw_Disc_Chk_A_H_Auto[1] OR Out_CYw_Disc_Chk_A_H_Auto[2]) AND AutoMode AND NOT Pause[1] AND NOT TimerQ_In_SenCY_Disc_Chk_A_H, PT := T#10s);
_e133(CLK := Output_A_Error_TON[23].Q);
IF _e133.Q THEN Output_A_Error_M[23] := TRUE; END_IF;
HMI_Message_Request[29] := _e133.Q;

